//------------------------------------------------------------------------------
// HMI : input registers (1001...), REAL = low word first
//------------------------------------------------------------------------------
	//--- ADM100W_1
	GVL_MODBUS.Input_register_TCP_HMI[1000] := GVL_COM.COM_ADM100W_1.HMI_OUTPUT_FREQUENCY.Word_value[0];                   // 1001 | ADM100W Frequency (low word)
	GVL_MODBUS.Input_register_TCP_HMI[1001] := GVL_COM.COM_ADM100W_1.HMI_OUTPUT_FREQUENCY.Word_value[1];                   // 1002 | ADM100W Frequency (high word)
	GVL_MODBUS.Input_register_TCP_HMI[1002] := GVL_COM.COM_ADM100W_1.HMI_OUTPUT_L1_L2_VOLTAGE.Word_value[0];               // 1003 | ADM100W L1-L2 Voltage (low word)
	GVL_MODBUS.Input_register_TCP_HMI[1003] := GVL_COM.COM_ADM100W_1.HMI_OUTPUT_L1_L2_VOLTAGE.Word_value[1];               // 1004 | ADM100W L1-L2 Voltage (high word)
	GVL_MODBUS.Input_register_TCP_HMI[1004] := GVL_COM.COM_ADM100W_1.HMI_OUTPUT_L1_N_VOLTAGE.Word_value[0];                // 1005 | ADM100W L1-N Voltage (low word)
	GVL_MODBUS.Input_register_TCP_HMI[1005] := GVL_COM.COM_ADM100W_1.HMI_OUTPUT_L1_N_VOLTAGE.Word_value[1];                // 1006 | ADM100W L1-N Voltage (high word)
	GVL_MODBUS.Input_register_TCP_HMI[1006] := GVL_COM.COM_ADM100W_1.HMI_OUTPUT_L1_CURRENT.Word_value[0];                  // 1007 | ADM100W L1 Current (low word)
	GVL_MODBUS.Input_register_TCP_HMI[1007] := GVL_COM.COM_ADM100W_1.HMI_OUTPUT_L1_CURRENT.Word_value[1];                  // 1008 | ADM100W L1 Current (high word)
	GVL_MODBUS.Input_register_TCP_HMI[1008] := GVL_COM.COM_ADM100W_1.HMI_OUTPUT_L1_ACTIVE_POWER.Word_value[0];             // 1009 | ADM100W L1 Active Power (low word)
	GVL_MODBUS.Input_register_TCP_HMI[1009] := GVL_COM.COM_ADM100W_1.HMI_OUTPUT_L1_ACTIVE_POWER.Word_value[1];             // 1010 | ADM100W L1 Active Power (high word)
	GVL_MODBUS.Input_register_TCP_HMI[1010] := GVL_COM.COM_ADM100W_1.HMI_OUTPUT_L1_APPARENT_POWER.Word_value[0];           // 1011 | ADM100W L1 Apparent Power (low word)
	GVL_MODBUS.Input_register_TCP_HMI[1011] := GVL_COM.COM_ADM100W_1.HMI_OUTPUT_L1_APPARENT_POWER.Word_value[1];           // 1012 | ADM100W L1 Apparent Power (high word)
	GVL_MODBUS.Input_register_TCP_HMI[1012] := GVL_COM.COM_ADM100W_1.HMI_OUTPUT_L1_REACTIVE_POWER.Word_value[0];           // 1013 | ADM100W L1 Reactive Power (low word)
	GVL_MODBUS.Input_register_TCP_HMI[1013] := GVL_COM.COM_ADM100W_1.HMI_OUTPUT_L1_REACTIVE_POWER.Word_value[1];           // 1014 | ADM100W L1 Reactive Power (high word)
	GVL_MODBUS.Input_register_TCP_HMI[1014] := GVL_COM.COM_ADM100W_1.HMI_OUTPUT_L1_CURRENT_PHASE_ANGLE.Word_value[0];      // 1015 | ADM100W L1 Current Phase Angle (low word)
	GVL_MODBUS.Input_register_TCP_HMI[1015] := GVL_COM.COM_ADM100W_1.HMI_OUTPUT_L1_CURRENT_PHASE_ANGLE.Word_value[1];      // 1016 | ADM100W L1 Current Phase Angle (high word)
	GVL_MODBUS.Input_register_TCP_HMI[1016] := GVL_COM.COM_ADM100W_1.HMI_OUTPUT_L1_POWER_FACTOR.Word_value[0];             // 1017 | ADM100W L1 Power Factor (low word)
	GVL_MODBUS.Input_register_TCP_HMI[1017] := GVL_COM.COM_ADM100W_1.HMI_OUTPUT_L1_POWER_FACTOR.Word_value[1];             // 1018 | ADM100W L1 Power Factor (high word)
	GVL_MODBUS.Input_register_TCP_HMI[1018] := GVL_COM.COM_ADM100W_1.HMI_OUTPUT_L1_VOLTAGE_THD.Word_value[0];              // 1019 | ADM100W L1 Voltage THD (low word)
	GVL_MODBUS.Input_register_TCP_HMI[1019] := GVL_COM.COM_ADM100W_1.HMI_OUTPUT_L1_VOLTAGE_THD.Word_value[1];              // 1020 | ADM100W L1 Voltage THD (high word)
	GVL_MODBUS.Input_register_TCP_HMI[1020] := GVL_COM.COM_ADM100W_1.HMI_OUTPUT_L1_CURRENT_THD.Word_value[0];              // 1021 | ADM100W L1 Current THD (low word)
	GVL_MODBUS.Input_register_TCP_HMI[1021] := GVL_COM.COM_ADM100W_1.HMI_OUTPUT_L1_CURRENT_THD.Word_value[1];              // 1022 | ADM100W L1 Current THD (high word)
	GVL_MODBUS.Input_register_TCP_HMI[1022] := GVL_COM.COM_ADM100W_1.HMI_OUTPUT_L1_MAX_LOAD.Word_value[0];                 // 1023 | ADM100W L1 Max Load (low word)
	GVL_MODBUS.Input_register_TCP_HMI[1023] := GVL_COM.COM_ADM100W_1.HMI_OUTPUT_L1_MAX_LOAD.Word_value[1];                 // 1024 | ADM100W L1 Max Load (high word)
	GVL_MODBUS.Input_register_TCP_HMI[1024] := GVL_COM.COM_ADM100W_1.HMI_OUTPUT_L1_L2_VOLTAGE_PHASE_ANGLE.Word_value[0];   // 1025 | ADM100W L1-L2 Voltage Phase Angle (low word)
	GVL_MODBUS.Input_register_TCP_HMI[1025] := GVL_COM.COM_ADM100W_1.HMI_OUTPUT_L1_L2_VOLTAGE_PHASE_ANGLE.Word_value[1];   // 1026 | ADM100W L1-L2 Voltage Phase Angle (high word)
	GVL_MODBUS.Input_register_TCP_HMI[1026] := GVL_COM.COM_ADM100W_1.HMI_OUTPUT_L2_L3_VOLTAGE.Word_value[0];               // 1027 | ADM100W L2-L3 Voltage (low word)
	GVL_MODBUS.Input_register_TCP_HMI[1027] := GVL_COM.COM_ADM100W_1.HMI_OUTPUT_L2_L3_VOLTAGE.Word_value[1];               // 1028 | ADM100W L2-L3 Voltage (high word)
	GVL_MODBUS.Input_register_TCP_HMI[1028] := GVL_COM.COM_ADM100W_1.HMI_OUTPUT_L2_N_VOLTAGE.Word_value[0];                // 1029 | ADM100W L2-N Voltage (low word)
	GVL_MODBUS.Input_register_TCP_HMI[1029] := GVL_COM.COM_ADM100W_1.HMI_OUTPUT_L2_N_VOLTAGE.Word_value[1];                // 1030 | ADM100W L2-N Voltage (high word)
	GVL_MODBUS.Input_register_TCP_HMI[1030] := GVL_COM.COM_ADM100W_1.HMI_OUTPUT_L2_CURRENT.Word_value[0];                  // 1031 | ADM100W L2 Current (low word)
	GVL_MODBUS.Input_register_TCP_HMI[1031] := GVL_COM.COM_ADM100W_1.HMI_OUTPUT_L2_CURRENT.Word_value[1];                  // 1032 | ADM100W L2 Current (high word)
	GVL_MODBUS.Input_register_TCP_HMI[1032] := GVL_COM.COM_ADM100W_1.HMI_OUTPUT_L2_ACTIVE_POWER.Word_value[0];             // 1033 | ADM100W L2 Active Power (low word)
	GVL_MODBUS.Input_register_TCP_HMI[1033] := GVL_COM.COM_ADM100W_1.HMI_OUTPUT_L2_ACTIVE_POWER.Word_value[1];             // 1034 | ADM100W L2 Active Power (high word)
	GVL_MODBUS.Input_register_TCP_HMI[1034] := GVL_COM.COM_ADM100W_1.HMI_OUTPUT_L2_APPARENT_POWER.Word_value[0];           // 1035 | ADM100W L2 Apparent Power (low word)
	GVL_MODBUS.Input_register_TCP_HMI[1035] := GVL_COM.COM_ADM100W_1.HMI_OUTPUT_L2_APPARENT_POWER.Word_value[1];           // 1036 | ADM100W L2 Apparent Power (high word)
	GVL_MODBUS.Input_register_TCP_HMI[1036] := GVL_COM.COM_ADM100W_1.HMI_OUTPUT_L2_REACTIVE_POWER.Word_value[0];           // 1037 | ADM100W L2 Reactive Power (low word)
	GVL_MODBUS.Input_register_TCP_HMI[1037] := GVL_COM.COM_ADM100W_1.HMI_OUTPUT_L2_REACTIVE_POWER.Word_value[1];           // 1038 | ADM100W L2 Reactive Power (high word)
	GVL_MODBUS.Input_register_TCP_HMI[1038] := GVL_COM.COM_ADM100W_1.HMI_OUTPUT_L2_CURRENT_PHASE_ANGLE.Word_value[0];      // 1039 | ADM100W L2 Current Phase Angle (low word)
	GVL_MODBUS.Input_register_TCP_HMI[1039] := GVL_COM.COM_ADM100W_1.HMI_OUTPUT_L2_CURRENT_PHASE_ANGLE.Word_value[1];      // 1040 | ADM100W L2 Current Phase Angle (high word)
	GVL_MODBUS.Input_register_TCP_HMI[1040] := GVL_COM.COM_ADM100W_1.HMI_OUTPUT_L2_POWER_FACTOR.Word_value[0];             // 1041 | ADM100W L2 Power Factor (low word)
	GVL_MODBUS.Input_register_TCP_HMI[1041] := GVL_COM.COM_ADM100W_1.HMI_OUTPUT_L2_POWER_FACTOR.Word_value[1];             // 1042 | ADM100W L2 Power Factor (high word)
	GVL_MODBUS.Input_register_TCP_HMI[1042] := GVL_COM.COM_ADM100W_1.HMI_OUTPUT_L2_VOLTAGE_THD.Word_value[0];              // 1043 | ADM100W L2 Voltage THD (low word)
	GVL_MODBUS.Input_register_TCP_HMI[1043] := GVL_COM.COM_ADM100W_1.HMI_OUTPUT_L2_VOLTAGE_THD.Word_value[1];              // 1044 | ADM100W L2 Voltage THD (high word)
	GVL_MODBUS.Input_register_TCP_HMI[1044] := GVL_COM.COM_ADM100W_1.HMI_OUTPUT_L2_CURRENT_THD.Word_value[0];              // 1045 | ADM100W L2 Current THD (low word)
	GVL_MODBUS.Input_register_TCP_HMI[1045] := GVL_COM.COM_ADM100W_1.HMI_OUTPUT_L2_CURRENT_THD.Word_value[1];              // 1046 | ADM100W L2 Current THD (high word)
	GVL_MODBUS.Input_register_TCP_HMI[1046] := GVL_COM.COM_ADM100W_1.HMI_OUTPUT_L2_MAX_LOAD.Word_value[0];                 // 1047 | ADM100W L2 Max Load (low word)
	GVL_MODBUS.Input_register_TCP_HMI[1047] := GVL_COM.COM_ADM100W_1.HMI_OUTPUT_L2_MAX_LOAD.Word_value[1];                 // 1048 | ADM100W L2 Max Load (high word)
	GVL_MODBUS.Input_register_TCP_HMI[1048] := GVL_COM.COM_ADM100W_1.HMI_OUTPUT_L1_L3_VOLTAGE_PHASE_ANGLE.Word_value[0];   // 1049 | ADM100W L1-L3 Voltage Phase Angle (low word)
	GVL_MODBUS.Input_register_TCP_HMI[1049] := GVL_COM.COM_ADM100W_1.HMI_OUTPUT_L1_L3_VOLTAGE_PHASE_ANGLE.Word_value[1];   // 1050 | ADM100W L1-L3 Voltage Phase Angle (high word)
	GVL_MODBUS.Input_register_TCP_HMI[1050] := GVL_COM.COM_ADM100W_1.HMI_OUTPUT_L3_L1_VOLTAGE.Word_value[0];               // 1051 | ADM100W L3-L1 Voltage (low word)
	GVL_MODBUS.Input_register_TCP_HMI[1051] := GVL_COM.COM_ADM100W_1.HMI_OUTPUT_L3_L1_VOLTAGE.Word_value[1];               // 1052 | ADM100W L3-L1 Voltage (high word)
	GVL_MODBUS.Input_register_TCP_HMI[1052] := GVL_COM.COM_ADM100W_1.HMI_OUTPUT_L3_N_VOLTAGE.Word_value[0];                // 1053 | ADM100W L3-N Voltage (low word)
	GVL_MODBUS.Input_register_TCP_HMI[1053] := GVL_COM.COM_ADM100W_1.HMI_OUTPUT_L3_N_VOLTAGE.Word_value[1];                // 1054 | ADM100W L3-N Voltage (high word)
	GVL_MODBUS.Input_register_TCP_HMI[1054] := GVL_COM.COM_ADM100W_1.HMI_OUTPUT_L3_CURRENT.Word_value[0];                  // 1055 | ADM100W L3 Current (low word)
	GVL_MODBUS.Input_register_TCP_HMI[1055] := GVL_COM.COM_ADM100W_1.HMI_OUTPUT_L3_CURRENT.Word_value[1];                  // 1056 | ADM100W L3 Current (high word)
	GVL_MODBUS.Input_register_TCP_HMI[1056] := GVL_COM.COM_ADM100W_1.HMI_OUTPUT_L3_ACTIVE_POWER.Word_value[0];             // 1057 | ADM100W L3 Active Power (low word)
	GVL_MODBUS.Input_register_TCP_HMI[1057] := GVL_COM.COM_ADM100W_1.HMI_OUTPUT_L3_ACTIVE_POWER.Word_value[1];             // 1058 | ADM100W L3 Active Power (high word)
	GVL_MODBUS.Input_register_TCP_HMI[1058] := GVL_COM.COM_ADM100W_1.HMI_OUTPUT_L3_APPARENT_POWER.Word_value[0];           // 1059 | ADM100W L3 Apparent Power (low word)
	GVL_MODBUS.Input_register_TCP_HMI[1059] := GVL_COM.COM_ADM100W_1.HMI_OUTPUT_L3_APPARENT_POWER.Word_value[1];           // 1060 | ADM100W L3 Apparent Power (high word)
	GVL_MODBUS.Input_register_TCP_HMI[1060] := GVL_COM.COM_ADM100W_1.HMI_OUTPUT_L3_REACTIVE_POWER.Word_value[0];           // 1061 | ADM100W L3 Reactive Power (low word)
	GVL_MODBUS.Input_register_TCP_HMI[1061] := GVL_COM.COM_ADM100W_1.HMI_OUTPUT_L3_REACTIVE_POWER.Word_value[1];           // 1062 | ADM100W L3 Reactive Power (high word)
	GVL_MODBUS.Input_register_TCP_HMI[1062] := GVL_COM.COM_ADM100W_1.HMI_OUTPUT_L3_CURRENT_PHASE_ANGLE.Word_value[0];      // 1063 | ADM100W L3 Current Phase Angle (low word)
	GVL_MODBUS.Input_register_TCP_HMI[1063] := GVL_COM.COM_ADM100W_1.HMI_OUTPUT_L3_CURRENT_PHASE_ANGLE.Word_value[1];      // 1064 | ADM100W L3 Current Phase Angle (high word)
	GVL_MODBUS.Input_register_TCP_HMI[1064] := GVL_COM.COM_ADM100W_1.HMI_OUTPUT_L3_POWER_FACTOR.Word_value[0];             // 1065 | ADM100W L3 Power Factor (low word)
	GVL_MODBUS.Input_register_TCP_HMI[1065] := GVL_COM.COM_ADM100W_1.HMI_OUTPUT_L3_POWER_FACTOR.Word_value[1];             // 1066 | ADM100W L3 Power Factor (high word)
	GVL_MODBUS.Input_register_TCP_HMI[1066] := GVL_COM.COM_ADM100W_1.HMI_OUTPUT_L3_VOLTAGE_THD.Word_value[0];              // 1067 | ADM100W L3 Voltage THD (low word)
	GVL_MODBUS.Input_register_TCP_HMI[1067] := GVL_COM.COM_ADM100W_1.HMI_OUTPUT_L3_VOLTAGE_THD.Word_value[1];              // 1068 | ADM100W L3 Voltage THD (high word)
	GVL_MODBUS.Input_register_TCP_HMI[1068] := GVL_COM.COM_ADM100W_1.HMI_OUTPUT_L3_CURRENT_THD.Word_value[0];              // 1069 | ADM100W L3 Current THD (low word)
	GVL_MODBUS.Input_register_TCP_HMI[1069] := GVL_COM.COM_ADM100W_1.HMI_OUTPUT_L3_CURRENT_THD.Word_value[1];              // 1070 | ADM100W L3 Current THD (high word)
	GVL_MODBUS.Input_register_TCP_HMI[1070] := GVL_COM.COM_ADM100W_1.HMI_OUTPUT_L3_MAX_LOAD.Word_value[0];                 // 1071 | ADM100W L3 Max Load (low word)
	GVL_MODBUS.Input_register_TCP_HMI[1071] := GVL_COM.COM_ADM100W_1.HMI_OUTPUT_L3_MAX_LOAD.Word_value[1];                 // 1072 | ADM100W L3 Max Load (high word)
	GVL_MODBUS.Input_register_TCP_HMI[1072] := GVL_COM.COM_ADM100W_1.HMI_OUTPUT_INTERNAL_TEMPERATURE.Word_value[0];        // 1073 | ADM100W Internal Temperature (low word)
	GVL_MODBUS.Input_register_TCP_HMI[1073] := GVL_COM.COM_ADM100W_1.HMI_OUTPUT_INTERNAL_TEMPERATURE.Word_value[1];        // 1074 | ADM100W Internal Temperature (high word)
	GVL_MODBUS.Input_register_TCP_HMI[1074] := GVL_COM.COM_ADM100W_1.HMI_OUTPUT_ACTIVE_ENERGY.Word_value[0];               // 1075 | ADM100W Active Energy (low word)
	GVL_MODBUS.Input_register_TCP_HMI[1075] := GVL_COM.COM_ADM100W_1.HMI_OUTPUT_ACTIVE_ENERGY.Word_value[1];               // 1076 | ADM100W Active Energy (high word)
	GVL_MODBUS.Input_register_TCP_HMI[1076] := GVL_COM.COM_ADM100W_1.HMI_OUTPUT_APPARENT_ENERGY.Word_value[0];             // 1077 | ADM100W Apparent Energy (low word)
	GVL_MODBUS.Input_register_TCP_HMI[1077] := GVL_COM.COM_ADM100W_1.HMI_OUTPUT_APPARENT_ENERGY.Word_value[1];             // 1078 | ADM100W Apparent Energy (high word)
	GVL_MODBUS.Input_register_TCP_HMI[1078] := GVL_COM.COM_ADM100W_1.HMI_OUTPUT_REACTIVE_ENERGY.Word_value[0];             // 1079 | ADM100W Reactive Energy (low word)
	GVL_MODBUS.Input_register_TCP_HMI[1079] := GVL_COM.COM_ADM100W_1.HMI_OUTPUT_REACTIVE_ENERGY.Word_value[1];             // 1080 | ADM100W Reactive Energy (high word)
	GVL_MODBUS.Input_register_TCP_HMI[1080] := GVL_COM.COM_ADM100W_1.HMI_OUTPUT_TOTAL_ACTIVE_POWER.Word_value[0];          // 1081 | ADM100W Total Active Power (low word)
	GVL_MODBUS.Input_register_TCP_HMI[1081] := GVL_COM.COM_ADM100W_1.HMI_OUTPUT_TOTAL_ACTIVE_POWER.Word_value[1];          // 1082 | ADM100W Total Active Power (high word)
	GVL_MODBUS.Input_register_TCP_HMI[1082] := GVL_COM.COM_ADM100W_1.HMI_OUTPUT_TOTAL_APPARENT_POWER.Word_value[0];        // 1083 | ADM100W Total Apparent Power (low word)
	GVL_MODBUS.Input_register_TCP_HMI[1083] := GVL_COM.COM_ADM100W_1.HMI_OUTPUT_TOTAL_APPARENT_POWER.Word_value[1];        // 1084 | ADM100W Total Apparent Power (high word)
	GVL_MODBUS.Input_register_TCP_HMI[1084] := GVL_COM.COM_ADM100W_1.HMI_OUTPUT_TOTAL_REACTIVE_POWER.Word_value[0];        // 1085 | ADM100W Total Reactive Power (low word)
	GVL_MODBUS.Input_register_TCP_HMI[1085] := GVL_COM.COM_ADM100W_1.HMI_OUTPUT_TOTAL_REACTIVE_POWER.Word_value[1];        // 1086 | ADM100W Total Reactive Power (high word)
	GVL_MODBUS.Input_register_TCP_HMI[1086] := GVL_COM.COM_ADM100W_1.HMI_OUTPUT_ALL_PHASE_POWER_FACTOR.Word_value[0];      // 1087 | ADM100W All Phase Power Factor (low word)
	GVL_MODBUS.Input_register_TCP_HMI[1087] := GVL_COM.COM_ADM100W_1.HMI_OUTPUT_ALL_PHASE_POWER_FACTOR.Word_value[1];      // 1088 | ADM100W All Phase Power Factor (high word)

	//--- DOSENSOR_1
	GVL_MODBUS.Input_register_TCP_HMI[1088] := GVL_COM.COM_DOSENSOR_1.HMI_OUTPUT_SIGNAL.Word_value[0];   // 1089 | DO Sensor Signal (low word)
	GVL_MODBUS.Input_register_TCP_HMI[1089] := GVL_COM.COM_DOSENSOR_1.HMI_OUTPUT_SIGNAL.Word_value[1];   // 1090 | DO Sensor Signal (high word)

	//--- DIP1500_1
	GVL_MODBUS.Input_register_TCP_HMI[1090] := GVL_COM.COM_DIP1500_1.HMI_OUTPUT_FIRMWARE_VERSION;                               // 1091 | DIP1500 Firmware Version
	GVL_MODBUS.Input_register_TCP_HMI[1091] := GVL_COM.COM_DIP1500_1.HMI_OUTPUT_HARDWARE_VERSION;                               // 1092 | DIP1500 Hardware Version
	GVL_MODBUS.Input_register_TCP_HMI[1092] := GVL_COM.COM_DIP1500_1.HMI_OUTPUT_TEMPERATURE;                                    // 1093 | DIP1500 Temperature
	GVL_MODBUS.Input_register_TCP_HMI[1093] := GVL_COM.COM_DIP1500_1.HMI_OUTPUT_FLOAT_LEVEL_ALARM;                              // 1094 | DIP1500 Float Level Alarm
	GVL_MODBUS.Input_register_TCP_HMI[1094] := GVL_COM.COM_DIP1500_1.HMI_OUTPUT_DIGITAL_OUTPUT_VALUE;                           // 1095 | DIP1500 Digital Output Value
	GVL_MODBUS.Input_register_TCP_HMI[1095] := GVL_COM.COM_DIP1500_1.HMI_OUTPUT_REAL_TIME_RUN_TIME_OR_VOLUME.Word_value[0];     // 1096 | DIP1500 Real-Time Run Time Or Volume (low word)
	GVL_MODBUS.Input_register_TCP_HMI[1096] := GVL_COM.COM_DIP1500_1.HMI_OUTPUT_REAL_TIME_RUN_TIME_OR_VOLUME.Word_value[1];     // 1097 | DIP1500 Real-Time Run Time Or Volume (high word)
	GVL_MODBUS.Input_register_TCP_HMI[1097] := GVL_COM.COM_DIP1500_1.HMI_OUTPUT_ACCUMULATED_RUN_TIME_OR_VOLUME.Word_value[0];   // 1098 | DIP1500 Accumulated Run Time Or Volume (low word)
	GVL_MODBUS.Input_register_TCP_HMI[1098] := GVL_COM.COM_DIP1500_1.HMI_OUTPUT_ACCUMULATED_RUN_TIME_OR_VOLUME.Word_value[1];   // 1099 | DIP1500 Accumulated Run Time Or Volume (high word)

GFC_COM_OUT := TRUE;

          
END_FUNCTION

FUNCTION GFC_EXC_IN : BOOL

            
//==============================================================================
// GFC_EXC_IN
// GVL_EXC -> GVL_EXC : functional units (UPI) to equipment, before GFB_INST
// Simple copies only, no conversion (conversions are done in the FBs)
//==============================================================================

//------------------------------------------------------------------------------
// Global local modes (UPI_LOCAL_FUXA, UPI_LOCAL_HMI, UPI_LOCAL_WEBVISU) to every equipment
//------------------------------------------------------------------------------
	//--- ADM100W_1
	GVL_EXC.EXC_ADM100W_1.UPI_INPUT_GLOBAL_LOCAL_FUXA := GVL_EXC.EXC_UPI_LOCAL_FUXA.UPI_OUTPUT_LOCAL_ACTIVE;
	GVL_EXC.EXC_ADM100W_1.UPI_INPUT_GLOBAL_LOCAL_HMI  := GVL_EXC.EXC_UPI_LOCAL_HMI.UPI_OUTPUT_LOCAL_ACTIVE;
	GVL_EXC.EXC_ADM100W_1.UPI_INPUT_GLOBAL_LOCAL_WEBVISU := GVL_EXC.EXC_UPI_LOCAL_WEBVISU.UPI_OUTPUT_LOCAL_ACTIVE;

	//--- DOSENSOR_1
	GVL_EXC.EXC_DOSENSOR_1.UPI_INPUT_GLOBAL_LOCAL_FUXA := GVL_EXC.EXC_UPI_LOCAL_FUXA.UPI_OUTPUT_LOCAL_ACTIVE;
	GVL_EXC.EXC_DOSENSOR_1.UPI_INPUT_GLOBAL_LOCAL_HMI  := GVL_EXC.EXC_UPI_LOCAL_HMI.UPI_OUTPUT_LOCAL_ACTIVE;
	GVL_EXC.EXC_DOSENSOR_1.UPI_INPUT_GLOBAL_LOCAL_WEBVISU := GVL_EXC.EXC_UPI_LOCAL_WEBVISU.UPI_OUTPUT_LOCAL_ACTIVE;

	//--- DIP1500_1
	GVL_EXC.EXC_DIP1500_1.UPI_INPUT_GLOBAL_LOCAL_FUXA := GVL_EXC.EXC_UPI_LOCAL_FUXA.UPI_OUTPUT_LOCAL_ACTIVE;
	GVL_EXC.EXC_DIP1500_1.UPI_INPUT_GLOBAL_LOCAL_HMI  := GVL_EXC.EXC_UPI_LOCAL_HMI.UPI_OUTPUT_LOCAL_ACTIVE;
	GVL_EXC.EXC_DIP1500_1.UPI_INPUT_GLOBAL_LOCAL_WEBVISU := GVL_EXC.EXC_UPI_LOCAL_WEBVISU.UPI_OUTPUT_LOCAL_ACTIVE;

GFC_EXC_IN := TRUE;

          
END_FUNCTION

FUNCTION GFC_EXC_OUT : BOOL

            
//==============================================================================
// GFC_EXC_OUT
// GVL_EXC -> GVL_EXC : equipment to equipment, after GFB_INST
// Simple copies only, no conversion (conversions are done in the FBs)
//==============================================================================

// Nothing to copy yet
GFC_EXC_OUT := TRUE;

          
END_FUNCTION

FUNCTION GFC_IO_IN : BOOL

            
//==============================================================================
// GFC_IO_IN
// GVL_IOMAP (PLC I/O cards) -> GVL_IO
// Simple copies only, no conversion (conversions are done in the FBs)
//==============================================================================

//------------------------------------------------------------------------------
// Digital inputs
//------------------------------------------------------------------------------
	//--- DOSENSOR_1
	GVL_IO.IO_DOSENSOR_1.INPUT_SENSOR_FAULT := GVL_IOMAP.IOMAP_DI_FAULT_DOSENSOR_1;


//------------------------------------------------------------------------------
// Analog inputs
//------------------------------------------------------------------------------
	//--- DOSENSOR_1
	GVL_IO.IO_DOSENSOR_1.INPUT_SIGNAL := GVL_IOMAP.IOMAP_AI_SIGNAL_DOSENSOR_1;

GFC_IO_IN := TRUE;

          
END_FUNCTION

FUNCTION GFC_IO_OUT : BOOL

            
//==============================================================================
// GFC_IO_OUT
// GVL_IO -> GVL_IOMAP (PLC I/O cards)
// Simple copies only, no conversion (conversions are done in the FBs)
//==============================================================================

//------------------------------------------------------------------------------
// Digital outputs
//------------------------------------------------------------------------------
	//--- DOSENSOR_1
	GVL_IOMAP.IOMAP_DO_HIGH_DOSENSOR_1 := GVL_IO.IO_DOSENSOR_1.OUTPUT_CALIBRATION_HIGH;
	GVL_IOMAP.IOMAP_DO_LOW_DOSENSOR_1  := GVL_IO.IO_DOSENSOR_1.OUTPUT_CALIBRATION_LOW;

GFC_IO_OUT := TRUE;

          
END_FUNCTION

FUNCTION_BLOCK FB_UPI_LOCAL_FUXA
  VAR_IN_OUT
    COM : DUT_COM_UPI_LOCAL_FUXA;  (* Requests and status with SCADA / HMI *)
    EXC : DUT_EXC_UPI_LOCAL_FUXA;  (* Status to equipment *)
  END_VAR
  VAR
    INTERN : DUT_INT_UPI_LOCAL_FUXA;  (* Internal variables *)
  END_VAR

            
//==============================================================================
// FB_UPI_LOCAL_FUXA
// Global FUXA local mode for every equipment
// Set by the FUXA local request, reset by the FUXA auto request (pulse or maintained, auto wins)
// The equipment read this status through GFC_EXC_IN and report their own local status themselves
//==============================================================================

//------------------------------------------------------------------------------
// 1. INPUTS
//------------------------------------------------------------------------------
	INTERN.LOCAL_REQUEST := COM.SCADA_INPUT_LOCAL_REQUEST;
	INTERN.AUTO_REQUEST  := COM.SCADA_INPUT_AUTO_REQUEST;


//------------------------------------------------------------------------------
// 2. PROCESSING
//------------------------------------------------------------------------------
	IF INTERN.LOCAL_REQUEST THEN
		INTERN.LOCAL_ACTIVE := TRUE;
	END_IF
	IF INTERN.AUTO_REQUEST THEN
		INTERN.LOCAL_ACTIVE := FALSE;
	END_IF


//------------------------------------------------------------------------------
// 3. OUTPUTS
//------------------------------------------------------------------------------
	//--- EXC : to every equipment (through GFC_EXC_IN)
	EXC.UPI_OUTPUT_LOCAL_ACTIVE := INTERN.LOCAL_ACTIVE;

	//--- COM : status
	COM.SCADA_OUTPUT_LOCAL_ACTIVE := INTERN.LOCAL_ACTIVE;


          
END_FUNCTION_BLOCK

FUNCTION_BLOCK FB_UPI_LOCAL_HMI
  VAR_IN_OUT
    COM : DUT_COM_UPI_LOCAL_HMI;  (* Requests and status with SCADA / HMI *)
    EXC : DUT_EXC_UPI_LOCAL_HMI;  (* Status to equipment *)
  END_VAR
  VAR
    INTERN : DUT_INT_UPI_LOCAL_HMI;  (* Internal variables *)
  END_VAR

            
//==============================================================================
// FB_UPI_LOCAL_HMI
// Global HMI local mode for every equipment
// Set by the HMI local request, reset by the HMI auto request (pulse or maintained, auto wins)
// The equipment read this status through GFC_EXC_IN and report their own local status themselves
//==============================================================================

//------------------------------------------------------------------------------
// 1. INPUTS
//------------------------------------------------------------------------------
	INTERN.LOCAL_REQUEST := COM.HMI_INPUT_LOCAL_REQUEST;
	INTERN.AUTO_REQUEST  := COM.HMI_INPUT_AUTO_REQUEST;


//------------------------------------------------------------------------------
// 2. PROCESSING
//------------------------------------------------------------------------------
	IF INTERN.LOCAL_REQUEST THEN
		INTERN.LOCAL_ACTIVE := TRUE;
	END_IF
	IF INTERN.AUTO_REQUEST THEN
		INTERN.LOCAL_ACTIVE := FALSE;
	END_IF


//------------------------------------------------------------------------------
// 3. OUTPUTS
//------------------------------------------------------------------------------
	//--- EXC : to every equipment (through GFC_EXC_IN)
	EXC.UPI_OUTPUT_LOCAL_ACTIVE := INTERN.LOCAL_ACTIVE;

	//--- COM : status
	COM.HMI_OUTPUT_LOCAL_ACTIVE   := INTERN.LOCAL_ACTIVE;
	COM.SCADA_OUTPUT_LOCAL_ACTIVE := INTERN.LOCAL_ACTIVE;   // also reported to FUXA


          
END_FUNCTION_BLOCK

FUNCTION_BLOCK GFB_INST
  VAR
    FB_ADM100W_1 : FB_INST_ADM100W;  (* Trumeter ADM100W power meter *)
    FB_DOSENSOR_1 : FB_INST_DOSENSOR;  (* Dissolved oxygen sensor *)
    FB_DIP1500_1 : FB_INST_DIP1500;  (* Kamoer DIP1500 peristaltic pump *)
  END_VAR

            
//==============================================================================
// GFB_INST
// Calls every equipment instance
// One block per equipment, all interfaces connected
//==============================================================================

//--- ADM100W_1 : Trumeter ADM100W power meter
FB_ADM100W_1(
	PA  := GVL_PA.PA_ADM100W_1,
	COM := GVL_COM.COM_ADM100W_1,
	EXC := GVL_EXC.EXC_ADM100W_1,
	IO  := GVL_IO.IO_ADM100W_1);

//--- DOSENSOR_1 : Dissolved oxygen sensor
FB_DOSENSOR_1(
	PA  := GVL_PA.PA_DOSENSOR_1,
	COM := GVL_COM.COM_DOSENSOR_1,
	EXC := GVL_EXC.EXC_DOSENSOR_1,
	IO  := GVL_IO.IO_DOSENSOR_1);

//--- DIP1500_1 : Kamoer DIP1500 peristaltic pump
FB_DIP1500_1(
	PA  := GVL_PA.PA_DIP1500_1,
	COM := GVL_COM.COM_DIP1500_1,
	EXC := GVL_EXC.EXC_DIP1500_1,
	IO  := GVL_IO.IO_DIP1500_1);

          
END_FUNCTION_BLOCK

FUNCTION_BLOCK GFB_UPI
  VAR
    FB_UPI_LOCAL_FUXA_1 : FB_UPI_LOCAL_FUXA;  (* Global FUXA local mode *)
    FB_UPI_LOCAL_HMI_1 : FB_UPI_LOCAL_HMI;  (* Global HMI local mode *)
    FB_UPI_LOCAL_WEBVISU_1 : FB_UPI_LOCAL_WEBVISU;  (* Global WEBVISU local mode *)
  END_VAR

            
//==============================================================================
// GFB_UPI
// Calls every functional unit (UPI)
// Runs before GFB_INST, results go to the equipment through GFC_EXC_IN
//==============================================================================

//--- UPI_LOCAL_FUXA : Global FUXA local mode
FB_UPI_LOCAL_FUXA_1(
	COM := GVL_COM.COM_UPI_LOCAL_FUXA,
	EXC := GVL_EXC.EXC_UPI_LOCAL_FUXA);

//--- UPI_LOCAL_HMI : Global HMI local mode
FB_UPI_LOCAL_HMI_1(
	COM := GVL_COM.COM_UPI_LOCAL_HMI,
	EXC := GVL_EXC.EXC_UPI_LOCAL_HMI);

//--- UPI_LOCAL_WEBVISU : Global WEBVISU local mode (direct IEC variables)
FB_UPI_LOCAL_WEBVISU_1(
	COM := GVL_COM.COM_UPI_LOCAL_WEBVISU,
	EXC := GVL_EXC.EXC_UPI_LOCAL_WEBVISU);

          
END_FUNCTION_BLOCK

FUNCTION_BLOCK FB_UPI_LOCAL_WEBVISU
  VAR_IN_OUT
    COM : DUT_COM_UPI_LOCAL_WEBVISU;  (* Direct IEC requests and status with WEBVISU *)
    EXC : DUT_EXC_UPI_LOCAL_WEBVISU;  (* Status to equipment *)
  END_VAR
  VAR
    INTERN : DUT_INT_UPI_LOCAL_WEBVISU;  (* Internal variables *)
  END_VAR

            
//==============================================================================
// FB_UPI_LOCAL_WEBVISU
// Global WEBVISU local mode for every equipment
// Set by the WEBVISU local request, reset by the WEBVISU auto request (pulse or maintained, auto wins)
// The equipment read this status through GFC_EXC_IN and report their own local status themselves
//==============================================================================

//------------------------------------------------------------------------------
// 1. INPUTS
//------------------------------------------------------------------------------
	INTERN.LOCAL_REQUEST := COM.WEBVISU_INPUT_LOCAL_REQUEST;
	INTERN.AUTO_REQUEST  := COM.WEBVISU_INPUT_AUTO_REQUEST;


//------------------------------------------------------------------------------
// 2. PROCESSING
//------------------------------------------------------------------------------
	IF INTERN.LOCAL_REQUEST THEN
		INTERN.LOCAL_ACTIVE := TRUE;
	END_IF
	IF INTERN.AUTO_REQUEST THEN
		INTERN.LOCAL_ACTIVE := FALSE;
	END_IF


//------------------------------------------------------------------------------
// 3. OUTPUTS
//------------------------------------------------------------------------------
	//--- EXC : to every equipment (through GFC_EXC_IN)
	EXC.UPI_OUTPUT_LOCAL_ACTIVE := INTERN.LOCAL_ACTIVE;

	//--- COM : status
	COM.WEBVISU_OUTPUT_LOCAL_ACTIVE := INTERN.LOCAL_ACTIVE;


          
END_FUNCTION_BLOCK

FUNCTION_BLOCK FB_INST_ADM100W
  VAR_IN_OUT
    PA : DUT_PA_ADM100W;  (* Parameters (persistent, GVL_PA) *)
    COM : DUT_COM_ADM100W;  (* Communication : Modbus RTU (COM_), SCADA FUXA (SCADA_), HMI (HMI_) *)
    EXC : DUT_EXC_ADM100W;  (* Exchanges : other equipment (EXC_), functional units (UPI_) *)
    IO : DUT_IO_ADM100W;  (* Wired PLC I/O *)
  END_VAR
  VAR
    INTERN : DUT_INT_ADM100W;  (* Internal variables *)
  END_VAR

            
//==============================================================================
// FB_INST_ADM100W
// Trumeter ADM100W power meter, Modbus RTU, 32-bit float MSW first (ABCD). No command : local mode is only reported
// 1. INPUTS     : requests, control mode, command source, equipment feedback -> INTERN
// 2. PROCESSING : on INTERN only
// 3. OUTPUTS    : INTERN -> COM / IO / EXC
// Control mode  : local WEBVISU > local HMI > local FUXA > auto (functional units)
//==============================================================================

//------------------------------------------------------------------------------
// 1. INPUTS
//------------------------------------------------------------------------------
	//--- Control mode requests (WEBVISU, HMI, FUXA, global UPI)
	INTERN.FUXA_LOCAL_REQUEST := COM.SCADA_INPUT_LOCAL_REQUEST;
	INTERN.FUXA_AUTO_REQUEST  := COM.SCADA_INPUT_AUTO_REQUEST;
	INTERN.HMI_LOCAL_REQUEST  := COM.HMI_INPUT_LOCAL_REQUEST;
	INTERN.HMI_AUTO_REQUEST   := COM.HMI_INPUT_AUTO_REQUEST;
	INTERN.GLOBAL_LOCAL_FUXA  := EXC.UPI_INPUT_GLOBAL_LOCAL_FUXA;
	INTERN.GLOBAL_LOCAL_HMI   := EXC.UPI_INPUT_GLOBAL_LOCAL_HMI;
	INTERN.WEBVISU_LOCAL_REQUEST := COM.WEBVISU_INPUT_LOCAL_REQUEST;
	INTERN.WEBVISU_AUTO_REQUEST  := COM.WEBVISU_INPUT_AUTO_REQUEST;
	INTERN.GLOBAL_LOCAL_WEBVISU  := EXC.UPI_INPUT_GLOBAL_LOCAL_WEBVISU;

	//--- Control mode
	// Individual memories : set by the local request, reset by the auto request (auto wins if both)
	IF INTERN.WEBVISU_LOCAL_REQUEST THEN
		INTERN.LOCAL_WEBVISU_INDIVIDUAL := TRUE;
	END_IF
	IF INTERN.WEBVISU_AUTO_REQUEST THEN
		INTERN.LOCAL_WEBVISU_INDIVIDUAL := FALSE;
	END_IF
	IF INTERN.HMI_LOCAL_REQUEST THEN
		INTERN.LOCAL_HMI_INDIVIDUAL := TRUE;
	END_IF
	IF INTERN.HMI_AUTO_REQUEST THEN
		INTERN.LOCAL_HMI_INDIVIDUAL := FALSE;
	END_IF
	IF INTERN.FUXA_LOCAL_REQUEST THEN
		INTERN.LOCAL_FUXA_INDIVIDUAL := TRUE;
	END_IF
	IF INTERN.FUXA_AUTO_REQUEST THEN
		INTERN.LOCAL_FUXA_INDIVIDUAL := FALSE;
	END_IF

	// Resulting mode : individual OR global, WEBVISU > HMI > FUXA > auto
	INTERN.LOCAL_WEBVISU := INTERN.LOCAL_WEBVISU_INDIVIDUAL OR INTERN.GLOBAL_LOCAL_WEBVISU;
	INTERN.LOCAL_HMI     := (INTERN.LOCAL_HMI_INDIVIDUAL OR INTERN.GLOBAL_LOCAL_HMI) AND NOT INTERN.LOCAL_WEBVISU;
	INTERN.LOCAL_FUXA    := (INTERN.LOCAL_FUXA_INDIVIDUAL OR INTERN.GLOBAL_LOCAL_FUXA) AND NOT INTERN.LOCAL_WEBVISU AND NOT INTERN.LOCAL_HMI;
	INTERN.AUTO          := NOT INTERN.LOCAL_WEBVISU AND NOT INTERN.LOCAL_HMI AND NOT INTERN.LOCAL_FUXA;

	//--- COM : alarms (coils 0..9)
	INTERN.ALARM_1  := COM.COM_INPUT_COILS[0].0;
	INTERN.ALARM_2  := COM.COM_INPUT_COILS[0].1;
	INTERN.ALARM_3  := COM.COM_INPUT_COILS[0].2;
	INTERN.ALARM_4  := COM.COM_INPUT_COILS[0].3;
	INTERN.ALARM_5  := COM.COM_INPUT_COILS[0].4;
	INTERN.ALARM_6  := COM.COM_INPUT_COILS[0].5;
	INTERN.ALARM_7  := COM.COM_INPUT_COILS[0].6;
	INTERN.ALARM_8  := COM.COM_INPUT_COILS[0].7;
	INTERN.ALARM_9  := COM.COM_INPUT_COILS[1].0;
	INTERN.ALARM_10 := COM.COM_INPUT_COILS[1].1;

	//--- COM : measures (input registers, MSW first)
	INTERN.FREQUENCY                 := FNC_WORDS_TO_REAL(High_word := COM.COM_INPUT_IR[0], Low_word := COM.COM_INPUT_IR[1]);
	INTERN.L1_L2_VOLTAGE             := FNC_WORDS_TO_REAL(High_word := COM.COM_INPUT_IR[2], Low_word := COM.COM_INPUT_IR[3]);
	INTERN.L1_N_VOLTAGE              := FNC_WORDS_TO_REAL(High_word := COM.COM_INPUT_IR[4], Low_word := COM.COM_INPUT_IR[5]);
	INTERN.L1_CURRENT                := FNC_WORDS_TO_REAL(High_word := COM.COM_INPUT_IR[6], Low_word := COM.COM_INPUT_IR[7]);
	INTERN.L1_ACTIVE_POWER           := FNC_WORDS_TO_REAL(High_word := COM.COM_INPUT_IR[8], Low_word := COM.COM_INPUT_IR[9]);
	INTERN.L1_APPARENT_POWER         := FNC_WORDS_TO_REAL(High_word := COM.COM_INPUT_IR[10], Low_word := COM.COM_INPUT_IR[11]);
	INTERN.L1_REACTIVE_POWER         := FNC_WORDS_TO_REAL(High_word := COM.COM_INPUT_IR[12], Low_word := COM.COM_INPUT_IR[13]);
	INTERN.L1_CURRENT_PHASE_ANGLE    := FNC_WORDS_TO_REAL(High_word := COM.COM_INPUT_IR[14], Low_word := COM.COM_INPUT_IR[15]);
	INTERN.L1_POWER_FACTOR           := FNC_WORDS_TO_REAL(High_word := COM.COM_INPUT_IR[16], Low_word := COM.COM_INPUT_IR[17]);
	INTERN.L1_VOLTAGE_THD            := FNC_WORDS_TO_REAL(High_word := COM.COM_INPUT_IR[18], Low_word := COM.COM_INPUT_IR[19]);
	INTERN.L1_CURRENT_THD            := FNC_WORDS_TO_REAL(High_word := COM.COM_INPUT_IR[20], Low_word := COM.COM_INPUT_IR[21]);
	INTERN.L1_MAX_LOAD               := FNC_WORDS_TO_REAL(High_word := COM.COM_INPUT_IR[22], Low_word := COM.COM_INPUT_IR[23]);
	INTERN.L1_L2_VOLTAGE_PHASE_ANGLE := FNC_WORDS_TO_REAL(High_word := COM.COM_INPUT_IR[24], Low_word := COM.COM_INPUT_IR[25]);
	INTERN.L2_L3_VOLTAGE             := FNC_WORDS_TO_REAL(High_word := COM.COM_INPUT_IR[26], Low_word := COM.COM_INPUT_IR[27]);
	INTERN.L2_N_VOLTAGE              := FNC_WORDS_TO_REAL(High_word := COM.COM_INPUT_IR[28], Low_word := COM.COM_INPUT_IR[29]);
	INTERN.L2_CURRENT                := FNC_WORDS_TO_REAL(High_word := COM.COM_INPUT_IR[30], Low_word := COM.COM_INPUT_IR[31]);
	INTERN.L2_ACTIVE_POWER           := FNC_WORDS_TO_REAL(High_word := COM.COM_INPUT_IR[32], Low_word := COM.COM_INPUT_IR[33]);
	INTERN.L2_APPARENT_POWER         := FNC_WORDS_TO_REAL(High_word := COM.COM_INPUT_IR[34], Low_word := COM.COM_INPUT_IR[35]);
	INTERN.L2_REACTIVE_POWER         := FNC_WORDS_TO_REAL(High_word := COM.COM_INPUT_IR[36], Low_word := COM.COM_INPUT_IR[37]);
	INTERN.L2_CURRENT_PHASE_ANGLE    := FNC_WORDS_TO_REAL(High_word := COM.COM_INPUT_IR[38], Low_word := COM.COM_INPUT_IR[39]);
	INTERN.L2_POWER_FACTOR           := FNC_WORDS_TO_REAL(High_word := COM.COM_INPUT_IR[40], Low_word := COM.COM_INPUT_IR[41]);
	INTERN.L2_VOLTAGE_THD            := FNC_WORDS_TO_REAL(High_word := COM.COM_INPUT_IR[42], Low_word := COM.COM_INPUT_IR[43]);
	INTERN.L2_CURRENT_THD            := FNC_WORDS_TO_REAL(High_word := COM.COM_INPUT_IR[44], Low_word := COM.COM_INPUT_IR[45]);
	INTERN.L2_MAX_LOAD               := FNC_WORDS_TO_REAL(High_word := COM.COM_INPUT_IR[46], Low_word := COM.COM_INPUT_IR[47]);
	INTERN.L1_L3_VOLTAGE_PHASE_ANGLE := FNC_WORDS_TO_REAL(High_word := COM.COM_INPUT_IR[48], Low_word := COM.COM_INPUT_IR[49]);
	INTERN.L3_L1_VOLTAGE             := FNC_WORDS_TO_REAL(High_word := COM.COM_INPUT_IR[50], Low_word := COM.COM_INPUT_IR[51]);
	INTERN.L3_N_VOLTAGE              := FNC_WORDS_TO_REAL(High_word := COM.COM_INPUT_IR[52], Low_word := COM.COM_INPUT_IR[53]);
	INTERN.L3_CURRENT                := FNC_WORDS_TO_REAL(High_word := COM.COM_INPUT_IR[54], Low_word := COM.COM_INPUT_IR[55]);
	INTERN.L3_ACTIVE_POWER           := FNC_WORDS_TO_REAL(High_word := COM.COM_INPUT_IR[56], Low_word := COM.COM_INPUT_IR[57]);
	INTERN.L3_APPARENT_POWER         := FNC_WORDS_TO_REAL(High_word := COM.COM_INPUT_IR[58], Low_word := COM.COM_INPUT_IR[59]);
	INTERN.L3_REACTIVE_POWER         := FNC_WORDS_TO_REAL(High_word := COM.COM_INPUT_IR[60], Low_word := COM.COM_INPUT_IR[61]);
	INTERN.L3_CURRENT_PHASE_ANGLE    := FNC_WORDS_TO_REAL(High_word := COM.COM_INPUT_IR[62], Low_word := COM.COM_INPUT_IR[63]);
	INTERN.L3_POWER_FACTOR           := FNC_WORDS_TO_REAL(High_word := COM.COM_INPUT_IR[64], Low_word := COM.COM_INPUT_IR[65]);
	INTERN.L3_VOLTAGE_THD            := FNC_WORDS_TO_REAL(High_word := COM.COM_INPUT_IR[66], Low_word := COM.COM_INPUT_IR[67]);
	INTERN.L3_CURRENT_THD            := FNC_WORDS_TO_REAL(High_word := COM.COM_INPUT_IR[68], Low_word := COM.COM_INPUT_IR[69]);
	INTERN.L3_MAX_LOAD               := FNC_WORDS_TO_REAL(High_word := COM.COM_INPUT_IR[70], Low_word := COM.COM_INPUT_IR[71]);
	INTERN.INTERNAL_TEMPERATURE      := FNC_WORDS_TO_REAL(High_word := COM.COM_INPUT_IR[72], Low_word := COM.COM_INPUT_IR[73]);
	INTERN.ACTIVE_ENERGY             := FNC_WORDS_TO_REAL(High_word := COM.COM_INPUT_IR[74], Low_word := COM.COM_INPUT_IR[75]);
	INTERN.APPARENT_ENERGY           := FNC_WORDS_TO_REAL(High_word := COM.COM_INPUT_IR[76], Low_word := COM.COM_INPUT_IR[77]);
	INTERN.REACTIVE_ENERGY           := FNC_WORDS_TO_REAL(High_word := COM.COM_INPUT_IR[78], Low_word := COM.COM_INPUT_IR[79]);
	INTERN.TOTAL_ACTIVE_POWER        := FNC_WORDS_TO_REAL(High_word := COM.COM_INPUT_IR[80], Low_word := COM.COM_INPUT_IR[81]);
	INTERN.TOTAL_APPARENT_POWER      := FNC_WORDS_TO_REAL(High_word := COM.COM_INPUT_IR[82], Low_word := COM.COM_INPUT_IR[83]);
	INTERN.TOTAL_REACTIVE_POWER      := FNC_WORDS_TO_REAL(High_word := COM.COM_INPUT_IR[84], Low_word := COM.COM_INPUT_IR[85]);
	INTERN.ALL_PHASE_POWER_FACTOR    := FNC_WORDS_TO_REAL(High_word := COM.COM_INPUT_IR[86], Low_word := COM.COM_INPUT_IR[87]);


//------------------------------------------------------------------------------
// 2. PROCESSING
//------------------------------------------------------------------------------
	// Nothing


//------------------------------------------------------------------------------
// 3. OUTPUTS
//------------------------------------------------------------------------------
	//--- COM : control mode status to SCADA, HMI and WEBVISU
	COM.SCADA_OUTPUT_LOCAL_FUXA_ACTIVE := INTERN.LOCAL_FUXA;
	COM.SCADA_OUTPUT_LOCAL_HMI_ACTIVE  := INTERN.LOCAL_HMI;
	COM.HMI_OUTPUT_LOCAL_ACTIVE        := INTERN.LOCAL_HMI;
	COM.WEBVISU_OUTPUT_LOCAL_ACTIVE        := INTERN.LOCAL_WEBVISU;
	COM.WEBVISU_OUTPUT_LOCAL_HMI_ACTIVE  := INTERN.LOCAL_HMI;
	COM.WEBVISU_OUTPUT_LOCAL_FUXA_ACTIVE := INTERN.LOCAL_FUXA;

	//--- EXC
	EXC.EXC_OUTPUT_FREQUENCY            := INTERN.FREQUENCY;
	EXC.EXC_OUTPUT_L1_N_VOLTAGE         := INTERN.L1_N_VOLTAGE;
	EXC.EXC_OUTPUT_L1_CURRENT           := INTERN.L1_CURRENT;
	EXC.EXC_OUTPUT_L1_ACTIVE_POWER      := INTERN.L1_ACTIVE_POWER;
	EXC.EXC_OUTPUT_L1_APPARENT_POWER    := INTERN.L1_APPARENT_POWER;
	EXC.EXC_OUTPUT_L1_REACTIVE_POWER    := INTERN.L1_REACTIVE_POWER;
	EXC.EXC_OUTPUT_L1_POWER_FACTOR      := INTERN.L1_POWER_FACTOR;
	EXC.EXC_OUTPUT_L1_VOLTAGE_THD       := INTERN.L1_VOLTAGE_THD;
	EXC.EXC_OUTPUT_L1_CURRENT_THD       := INTERN.L1_CURRENT_THD;
	EXC.EXC_OUTPUT_L1_MAX_LOAD          := INTERN.L1_MAX_LOAD;
	EXC.EXC_OUTPUT_INTERNAL_TEMPERATURE := INTERN.INTERNAL_TEMPERATURE;
	EXC.EXC_OUTPUT_ACTIVE_ENERGY        := INTERN.ACTIVE_ENERGY;
	// EXC.EXC_OUTPUT_DATA_VALID : not managed yet (no Modbus diagnostic)

	//--- COM : alarms to SCADA, HMI and WEBVISU
	COM.SCADA_OUTPUT_ALARM_1_STATUS  := INTERN.ALARM_1;
	COM.HMI_OUTPUT_ALARM_1_STATUS    := INTERN.ALARM_1;
	COM.WEBVISU_OUTPUT_ALARM_1_STATUS    := INTERN.ALARM_1;
	COM.SCADA_OUTPUT_ALARM_2_STATUS  := INTERN.ALARM_2;
	COM.HMI_OUTPUT_ALARM_2_STATUS    := INTERN.ALARM_2;
	COM.WEBVISU_OUTPUT_ALARM_2_STATUS    := INTERN.ALARM_2;
	COM.SCADA_OUTPUT_ALARM_3_STATUS  := INTERN.ALARM_3;
	COM.HMI_OUTPUT_ALARM_3_STATUS    := INTERN.ALARM_3;
	COM.WEBVISU_OUTPUT_ALARM_3_STATUS    := INTERN.ALARM_3;
	COM.SCADA_OUTPUT_ALARM_4_STATUS  := INTERN.ALARM_4;
	COM.HMI_OUTPUT_ALARM_4_STATUS    := INTERN.ALARM_4;
	COM.WEBVISU_OUTPUT_ALARM_4_STATUS    := INTERN.ALARM_4;
	COM.SCADA_OUTPUT_ALARM_5_STATUS  := INTERN.ALARM_5;
	COM.HMI_OUTPUT_ALARM_5_STATUS    := INTERN.ALARM_5;
	COM.WEBVISU_OUTPUT_ALARM_5_STATUS    := INTERN.ALARM_5;
	COM.SCADA_OUTPUT_ALARM_6_STATUS  := INTERN.ALARM_6;
	COM.HMI_OUTPUT_ALARM_6_STATUS    := INTERN.ALARM_6;
	COM.WEBVISU_OUTPUT_ALARM_6_STATUS    := INTERN.ALARM_6;
	COM.SCADA_OUTPUT_ALARM_7_STATUS  := INTERN.ALARM_7;
	COM.HMI_OUTPUT_ALARM_7_STATUS    := INTERN.ALARM_7;
	COM.WEBVISU_OUTPUT_ALARM_7_STATUS    := INTERN.ALARM_7;
	COM.SCADA_OUTPUT_ALARM_8_STATUS  := INTERN.ALARM_8;
	COM.HMI_OUTPUT_ALARM_8_STATUS    := INTERN.ALARM_8;
	COM.WEBVISU_OUTPUT_ALARM_8_STATUS    := INTERN.ALARM_8;
	COM.SCADA_OUTPUT_ALARM_9_STATUS  := INTERN.ALARM_9;
	COM.HMI_OUTPUT_ALARM_9_STATUS    := INTERN.ALARM_9;
	COM.WEBVISU_OUTPUT_ALARM_9_STATUS    := INTERN.ALARM_9;
	COM.SCADA_OUTPUT_ALARM_10_STATUS := INTERN.ALARM_10;
	COM.HMI_OUTPUT_ALARM_10_STATUS   := INTERN.ALARM_10;
	COM.WEBVISU_OUTPUT_ALARM_10_STATUS   := INTERN.ALARM_10;

	//--- COM : measures to SCADA, HMI and WEBVISU
	COM.SCADA_OUTPUT_FREQUENCY.Real_value                 := INTERN.FREQUENCY;
	COM.HMI_OUTPUT_FREQUENCY.Real_value                   := INTERN.FREQUENCY;
	COM.WEBVISU_OUTPUT_FREQUENCY.Real_value                   := INTERN.FREQUENCY;
	COM.SCADA_OUTPUT_L1_L2_VOLTAGE.Real_value             := INTERN.L1_L2_VOLTAGE;
	COM.HMI_OUTPUT_L1_L2_VOLTAGE.Real_value               := INTERN.L1_L2_VOLTAGE;
	COM.WEBVISU_OUTPUT_L1_L2_VOLTAGE.Real_value               := INTERN.L1_L2_VOLTAGE;
	COM.SCADA_OUTPUT_L1_N_VOLTAGE.Real_value              := INTERN.L1_N_VOLTAGE;
	COM.HMI_OUTPUT_L1_N_VOLTAGE.Real_value                := INTERN.L1_N_VOLTAGE;
	COM.WEBVISU_OUTPUT_L1_N_VOLTAGE.Real_value                := INTERN.L1_N_VOLTAGE;
	COM.SCADA_OUTPUT_L1_CURRENT.Real_value                := INTERN.L1_CURRENT;
	COM.HMI_OUTPUT_L1_CURRENT.Real_value                  := INTERN.L1_CURRENT;
	COM.WEBVISU_OUTPUT_L1_CURRENT.Real_value                  := INTERN.L1_CURRENT;
	COM.SCADA_OUTPUT_L1_ACTIVE_POWER.Real_value           := INTERN.L1_ACTIVE_POWER;
	COM.HMI_OUTPUT_L1_ACTIVE_POWER.Real_value             := INTERN.L1_ACTIVE_POWER;
	COM.WEBVISU_OUTPUT_L1_ACTIVE_POWER.Real_value             := INTERN.L1_ACTIVE_POWER;
	COM.SCADA_OUTPUT_L1_APPARENT_POWER.Real_value         := INTERN.L1_APPARENT_POWER;
	COM.HMI_OUTPUT_L1_APPARENT_POWER.Real_value           := INTERN.L1_APPARENT_POWER;
	COM.WEBVISU_OUTPUT_L1_APPARENT_POWER.Real_value           := INTERN.L1_APPARENT_POWER;
	COM.SCADA_OUTPUT_L1_REACTIVE_POWER.Real_value         := INTERN.L1_REACTIVE_POWER;
	COM.HMI_OUTPUT_L1_REACTIVE_POWER.Real_value           := INTERN.L1_REACTIVE_POWER;
	COM.WEBVISU_OUTPUT_L1_REACTIVE_POWER.Real_value           := INTERN.L1_REACTIVE_POWER;
	COM.SCADA_OUTPUT_L1_CURRENT_PHASE_ANGLE.Real_value    := INTERN.L1_CURRENT_PHASE_ANGLE;
	COM.HMI_OUTPUT_L1_CURRENT_PHASE_ANGLE.Real_value      := INTERN.L1_CURRENT_PHASE_ANGLE;
	COM.WEBVISU_OUTPUT_L1_CURRENT_PHASE_ANGLE.Real_value      := INTERN.L1_CURRENT_PHASE_ANGLE;
	COM.SCADA_OUTPUT_L1_POWER_FACTOR.Real_value           := INTERN.L1_POWER_FACTOR;
	COM.HMI_OUTPUT_L1_POWER_FACTOR.Real_value             := INTERN.L1_POWER_FACTOR;
	COM.WEBVISU_OUTPUT_L1_POWER_FACTOR.Real_value             := INTERN.L1_POWER_FACTOR;
	COM.SCADA_OUTPUT_L1_VOLTAGE_THD.Real_value            := INTERN.L1_VOLTAGE_THD;
	COM.HMI_OUTPUT_L1_VOLTAGE_THD.Real_value              := INTERN.L1_VOLTAGE_THD;
	COM.WEBVISU_OUTPUT_L1_VOLTAGE_THD.Real_value              := INTERN.L1_VOLTAGE_THD;
	COM.SCADA_OUTPUT_L1_CURRENT_THD.Real_value            := INTERN.L1_CURRENT_THD;
	COM.HMI_OUTPUT_L1_CURRENT_THD.Real_value              := INTERN.L1_CURRENT_THD;
	COM.WEBVISU_OUTPUT_L1_CURRENT_THD.Real_value              := INTERN.L1_CURRENT_THD;
	COM.SCADA_OUTPUT_L1_MAX_LOAD.Real_value               := INTERN.L1_MAX_LOAD;
	COM.HMI_OUTPUT_L1_MAX_LOAD.Real_value                 := INTERN.L1_MAX_LOAD;
	COM.WEBVISU_OUTPUT_L1_MAX_LOAD.Real_value                 := INTERN.L1_MAX_LOAD;
	COM.SCADA_OUTPUT_L1_L2_VOLTAGE_PHASE_ANGLE.Real_value := INTERN.L1_L2_VOLTAGE_PHASE_ANGLE;
	COM.HMI_OUTPUT_L1_L2_VOLTAGE_PHASE_ANGLE.Real_value   := INTERN.L1_L2_VOLTAGE_PHASE_ANGLE;
	COM.WEBVISU_OUTPUT_L1_L2_VOLTAGE_PHASE_ANGLE.Real_value   := INTERN.L1_L2_VOLTAGE_PHASE_ANGLE;
	COM.SCADA_OUTPUT_L2_L3_VOLTAGE.Real_value             := INTERN.L2_L3_VOLTAGE;
	COM.HMI_OUTPUT_L2_L3_VOLTAGE.Real_value               := INTERN.L2_L3_VOLTAGE;
	COM.WEBVISU_OUTPUT_L2_L3_VOLTAGE.Real_value               := INTERN.L2_L3_VOLTAGE;
	COM.SCADA_OUTPUT_L2_N_VOLTAGE.Real_value              := INTERN.L2_N_VOLTAGE;
	COM.HMI_OUTPUT_L2_N_VOLTAGE.Real_value                := INTERN.L2_N_VOLTAGE;
	COM.WEBVISU_OUTPUT_L2_N_VOLTAGE.Real_value                := INTERN.L2_N_VOLTAGE;
	COM.SCADA_OUTPUT_L2_CURRENT.Real_value                := INTERN.L2_CURRENT;
	COM.HMI_OUTPUT_L2_CURRENT.Real_value                  := INTERN.L2_CURRENT;
	COM.WEBVISU_OUTPUT_L2_CURRENT.Real_value                  := INTERN.L2_CURRENT;
	COM.SCADA_OUTPUT_L2_ACTIVE_POWER.Real_value           := INTERN.L2_ACTIVE_POWER;
	COM.HMI_OUTPUT_L2_ACTIVE_POWER.Real_value             := INTERN.L2_ACTIVE_POWER;
	COM.WEBVISU_OUTPUT_L2_ACTIVE_POWER.Real_value             := INTERN.L2_ACTIVE_POWER;
	COM.SCADA_OUTPUT_L2_APPARENT_POWER.Real_value         := INTERN.L2_APPARENT_POWER;
	COM.HMI_OUTPUT_L2_APPARENT_POWER.Real_value           := INTERN.L2_APPARENT_POWER;
	COM.WEBVISU_OUTPUT_L2_APPARENT_POWER.Real_value           := INTERN.L2_APPARENT_POWER;
	COM.SCADA_OUTPUT_L2_REACTIVE_POWER.Real_value         := INTERN.L2_REACTIVE_POWER;
	COM.HMI_OUTPUT_L2_REACTIVE_POWER.Real_value           := INTERN.L2_REACTIVE_POWER;
	COM.WEBVISU_OUTPUT_L2_REACTIVE_POWER.Real_value           := INTERN.L2_REACTIVE_POWER;
	COM.SCADA_OUTPUT_L2_CURRENT_PHASE_ANGLE.Real_value    := INTERN.L2_CURRENT_PHASE_ANGLE;
	COM.HMI_OUTPUT_L2_CURRENT_PHASE_ANGLE.Real_value      := INTERN.L2_CURRENT_PHASE_ANGLE;
	COM.WEBVISU_OUTPUT_L2_CURRENT_PHASE_ANGLE.Real_value      := INTERN.L2_CURRENT_PHASE_ANGLE;
	COM.SCADA_OUTPUT_L2_POWER_FACTOR.Real_value           := INTERN.L2_POWER_FACTOR;
	COM.HMI_OUTPUT_L2_POWER_FACTOR.Real_value             := INTERN.L2_POWER_FACTOR;
	COM.WEBVISU_OUTPUT_L2_POWER_FACTOR.Real_value             := INTERN.L2_POWER_FACTOR;
	COM.SCADA_OUTPUT_L2_VOLTAGE_THD.Real_value            := INTERN.L2_VOLTAGE_THD;
	COM.HMI_OUTPUT_L2_VOLTAGE_THD.Real_value              := INTERN.L2_VOLTAGE_THD;
	COM.WEBVISU_OUTPUT_L2_VOLTAGE_THD.Real_value              := INTERN.L2_VOLTAGE_THD;
	COM.SCADA_OUTPUT_L2_CURRENT_THD.Real_value            := INTERN.L2_CURRENT_THD;
	COM.HMI_OUTPUT_L2_CURRENT_THD.Real_value              := INTERN.L2_CURRENT_THD;
	COM.WEBVISU_OUTPUT_L2_CURRENT_THD.Real_value              := INTERN.L2_CURRENT_THD;
	COM.SCADA_OUTPUT_L2_MAX_LOAD.Real_value               := INTERN.L2_MAX_LOAD;
	COM.HMI_OUTPUT_L2_MAX_LOAD.Real_value                 := INTERN.L2_MAX_LOAD;
	COM.WEBVISU_OUTPUT_L2_MAX_LOAD.Real_value                 := INTERN.L2_MAX_LOAD;
	COM.SCADA_OUTPUT_L1_L3_VOLTAGE_PHASE_ANGLE.Real_value := INTERN.L1_L3_VOLTAGE_PHASE_ANGLE;
	COM.HMI_OUTPUT_L1_L3_VOLTAGE_PHASE_ANGLE.Real_value   := INTERN.L1_L3_VOLTAGE_PHASE_ANGLE;
	COM.WEBVISU_OUTPUT_L1_L3_VOLTAGE_PHASE_ANGLE.Real_value   := INTERN.L1_L3_VOLTAGE_PHASE_ANGLE;
	COM.SCADA_OUTPUT_L3_L1_VOLTAGE.Real_value             := INTERN.L3_L1_VOLTAGE;
	COM.HMI_OUTPUT_L3_L1_VOLTAGE.Real_value               := INTERN.L3_L1_VOLTAGE;
	COM.WEBVISU_OUTPUT_L3_L1_VOLTAGE.Real_value               := INTERN.L3_L1_VOLTAGE;
	COM.SCADA_OUTPUT_L3_N_VOLTAGE.Real_value              := INTERN.L3_N_VOLTAGE;
	COM.HMI_OUTPUT_L3_N_VOLTAGE.Real_value                := INTERN.L3_N_VOLTAGE;
	COM.WEBVISU_OUTPUT_L3_N_VOLTAGE.Real_value                := INTERN.L3_N_VOLTAGE;
	COM.SCADA_OUTPUT_L3_CURRENT.Real_value                := INTERN.L3_CURRENT;
	COM.HMI_OUTPUT_L3_CURRENT.Real_value                  := INTERN.L3_CURRENT;
	COM.WEBVISU_OUTPUT_L3_CURRENT.Real_value                  := INTERN.L3_CURRENT;
	COM.SCADA_OUTPUT_L3_ACTIVE_POWER.Real_value           := INTERN.L3_ACTIVE_POWER;
	COM.HMI_OUTPUT_L3_ACTIVE_POWER.Real_value             := INTERN.L3_ACTIVE_POWER;
	COM.WEBVISU_OUTPUT_L3_ACTIVE_POWER.Real_value             := INTERN.L3_ACTIVE_POWER;
	COM.SCADA_OUTPUT_L3_APPARENT_POWER.Real_value         := INTERN.L3_APPARENT_POWER;
	COM.HMI_OUTPUT_L3_APPARENT_POWER.Real_value           := INTERN.L3_APPARENT_POWER;
	COM.WEBVISU_OUTPUT_L3_APPARENT_POWER.Real_value           := INTERN.L3_APPARENT_POWER;
	COM.SCADA_OUTPUT_L3_REACTIVE_POWER.Real_value         := INTERN.L3_REACTIVE_POWER;
	COM.HMI_OUTPUT_L3_REACTIVE_POWER.Real_value           := INTERN.L3_REACTIVE_POWER;
	COM.WEBVISU_OUTPUT_L3_REACTIVE_POWER.Real_value           := INTERN.L3_REACTIVE_POWER;
	COM.SCADA_OUTPUT_L3_CURRENT_PHASE_ANGLE.Real_value    := INTERN.L3_CURRENT_PHASE_ANGLE;
	COM.HMI_OUTPUT_L3_CURRENT_PHASE_ANGLE.Real_value      := INTERN.L3_CURRENT_PHASE_ANGLE;
	COM.WEBVISU_OUTPUT_L3_CURRENT_PHASE_ANGLE.Real_value      := INTERN.L3_CURRENT_PHASE_ANGLE;
	COM.SCADA_OUTPUT_L3_POWER_FACTOR.Real_value           := INTERN.L3_POWER_FACTOR;
	COM.HMI_OUTPUT_L3_POWER_FACTOR.Real_value             := INTERN.L3_POWER_FACTOR;
	COM.WEBVISU_OUTPUT_L3_POWER_FACTOR.Real_value             := INTERN.L3_POWER_FACTOR;
	COM.SCADA_OUTPUT_L3_VOLTAGE_THD.Real_value            := INTERN.L3_VOLTAGE_THD;
	COM.HMI_OUTPUT_L3_VOLTAGE_THD.Real_value              := INTERN.L3_VOLTAGE_THD;
	COM.WEBVISU_OUTPUT_L3_VOLTAGE_THD.Real_value              := INTERN.L3_VOLTAGE_THD;
	COM.SCADA_OUTPUT_L3_CURRENT_THD.Real_value            := INTERN.L3_CURRENT_THD;
	COM.HMI_OUTPUT_L3_CURRENT_THD.Real_value              := INTERN.L3_CURRENT_THD;
	COM.WEBVISU_OUTPUT_L3_CURRENT_THD.Real_value              := INTERN.L3_CURRENT_THD;
	COM.SCADA_OUTPUT_L3_MAX_LOAD.Real_value               := INTERN.L3_MAX_LOAD;
	COM.HMI_OUTPUT_L3_MAX_LOAD.Real_value                 := INTERN.L3_MAX_LOAD;
	COM.WEBVISU_OUTPUT_L3_MAX_LOAD.Real_value                 := INTERN.L3_MAX_LOAD;
	COM.SCADA_OUTPUT_INTERNAL_TEMPERATURE.Real_value      := INTERN.INTERNAL_TEMPERATURE;
	COM.HMI_OUTPUT_INTERNAL_TEMPERATURE.Real_value        := INTERN.INTERNAL_TEMPERATURE;
	COM.WEBVISU_OUTPUT_INTERNAL_TEMPERATURE.Real_value        := INTERN.INTERNAL_TEMPERATURE;
	COM.SCADA_OUTPUT_ACTIVE_ENERGY.Real_value             := INTERN.ACTIVE_ENERGY;
	COM.HMI_OUTPUT_ACTIVE_ENERGY.Real_value               := INTERN.ACTIVE_ENERGY;
	COM.WEBVISU_OUTPUT_ACTIVE_ENERGY.Real_value               := INTERN.ACTIVE_ENERGY;
	COM.SCADA_OUTPUT_APPARENT_ENERGY.Real_value           := INTERN.APPARENT_ENERGY;
	COM.HMI_OUTPUT_APPARENT_ENERGY.Real_value             := INTERN.APPARENT_ENERGY;
	COM.WEBVISU_OUTPUT_APPARENT_ENERGY.Real_value             := INTERN.APPARENT_ENERGY;
	COM.SCADA_OUTPUT_REACTIVE_ENERGY.Real_value           := INTERN.REACTIVE_ENERGY;
	COM.HMI_OUTPUT_REACTIVE_ENERGY.Real_value             := INTERN.REACTIVE_ENERGY;
	COM.WEBVISU_OUTPUT_REACTIVE_ENERGY.Real_value             := INTERN.REACTIVE_ENERGY;
	COM.SCADA_OUTPUT_TOTAL_ACTIVE_POWER.Real_value        := INTERN.TOTAL_ACTIVE_POWER;
	COM.HMI_OUTPUT_TOTAL_ACTIVE_POWER.Real_value          := INTERN.TOTAL_ACTIVE_POWER;
	COM.WEBVISU_OUTPUT_TOTAL_ACTIVE_POWER.Real_value          := INTERN.TOTAL_ACTIVE_POWER;
	COM.SCADA_OUTPUT_TOTAL_APPARENT_POWER.Real_value      := INTERN.TOTAL_APPARENT_POWER;
	COM.HMI_OUTPUT_TOTAL_APPARENT_POWER.Real_value        := INTERN.TOTAL_APPARENT_POWER;
	COM.WEBVISU_OUTPUT_TOTAL_APPARENT_POWER.Real_value        := INTERN.TOTAL_APPARENT_POWER;
	COM.SCADA_OUTPUT_TOTAL_REACTIVE_POWER.Real_value      := INTERN.TOTAL_REACTIVE_POWER;
	COM.HMI_OUTPUT_TOTAL_REACTIVE_POWER.Real_value        := INTERN.TOTAL_REACTIVE_POWER;
	COM.WEBVISU_OUTPUT_TOTAL_REACTIVE_POWER.Real_value        := INTERN.TOTAL_REACTIVE_POWER;
	COM.SCADA_OUTPUT_ALL_PHASE_POWER_FACTOR.Real_value    := INTERN.ALL_PHASE_POWER_FACTOR;
	COM.HMI_OUTPUT_ALL_PHASE_POWER_FACTOR.Real_value      := INTERN.ALL_PHASE_POWER_FACTOR;
	COM.WEBVISU_OUTPUT_ALL_PHASE_POWER_FACTOR.Real_value      := INTERN.ALL_PHASE_POWER_FACTOR;


          
END_FUNCTION_BLOCK

FUNCTION_BLOCK FB_INST_DIP1500
  VAR_IN_OUT
    PA : DUT_PA_DIP1500;  (* Parameters (persistent, GVL_PA) *)
    COM : DUT_COM_DIP1500;  (* Communication : Modbus RTU (COM_), SCADA FUXA (SCADA_), HMI (HMI_) *)
    EXC : DUT_EXC_DIP1500;  (* Exchanges : other equipment (EXC_), functional units (UPI_) *)
    IO : DUT_IO_DIP1500;  (* Wired PLC I/O *)
  END_VAR
  VAR
    INTERN : DUT_INT_DIP1500;  (* Internal variables *)
    TON_PULSE : TON;  (* Square wave timer *)
    TOF_CMD_WINDOW : TOF;  (* Command write window *)
    R_TRIG_FLASH : R_TRIG;  (* Flash save request edge *)
    TP_FLASH : TP;  (* Flash save pulse *)
  END_VAR

            
//==============================================================================
// FB_INST_DIP1500
// Kamoer DIP1500 peristaltic pump, Modbus RTU, 32-bit low word first (CDAB)
// 1. INPUTS     : requests, control mode, command source, equipment feedback -> INTERN
// 2. PROCESSING : on INTERN only
// 3. OUTPUTS    : INTERN -> COM / IO / EXC
// Parameters    : pump configuration in PA (persistent), changed from the active local supervision
// Control mode  : local WEBVISU > local HMI > local FUXA > auto (functional units)
//==============================================================================

//------------------------------------------------------------------------------
// 1. INPUTS
//------------------------------------------------------------------------------
	//--- Control mode requests (WEBVISU, HMI, FUXA, global UPI)
	INTERN.FUXA_LOCAL_REQUEST := COM.SCADA_INPUT_LOCAL_REQUEST;
	INTERN.FUXA_AUTO_REQUEST  := COM.SCADA_INPUT_AUTO_REQUEST;
	INTERN.HMI_LOCAL_REQUEST  := COM.HMI_INPUT_LOCAL_REQUEST;
	INTERN.HMI_AUTO_REQUEST   := COM.HMI_INPUT_AUTO_REQUEST;
	INTERN.GLOBAL_LOCAL_FUXA  := EXC.UPI_INPUT_GLOBAL_LOCAL_FUXA;
	INTERN.GLOBAL_LOCAL_HMI   := EXC.UPI_INPUT_GLOBAL_LOCAL_HMI;
	INTERN.WEBVISU_LOCAL_REQUEST := COM.WEBVISU_INPUT_LOCAL_REQUEST;
	INTERN.WEBVISU_AUTO_REQUEST  := COM.WEBVISU_INPUT_AUTO_REQUEST;
	INTERN.GLOBAL_LOCAL_WEBVISU  := EXC.UPI_INPUT_GLOBAL_LOCAL_WEBVISU;

	//--- Control mode
	// Individual memories : set by the local request, reset by the auto request (auto wins if both)
	IF INTERN.WEBVISU_LOCAL_REQUEST THEN
		INTERN.LOCAL_WEBVISU_INDIVIDUAL := TRUE;
	END_IF
	IF INTERN.WEBVISU_AUTO_REQUEST THEN
		INTERN.LOCAL_WEBVISU_INDIVIDUAL := FALSE;
	END_IF
	IF INTERN.HMI_LOCAL_REQUEST THEN
		INTERN.LOCAL_HMI_INDIVIDUAL := TRUE;
	END_IF
	IF INTERN.HMI_AUTO_REQUEST THEN
		INTERN.LOCAL_HMI_INDIVIDUAL := FALSE;
	END_IF
	IF INTERN.FUXA_LOCAL_REQUEST THEN
		INTERN.LOCAL_FUXA_INDIVIDUAL := TRUE;
	END_IF
	IF INTERN.FUXA_AUTO_REQUEST THEN
		INTERN.LOCAL_FUXA_INDIVIDUAL := FALSE;
	END_IF

	// Resulting mode : individual OR global, WEBVISU > HMI > FUXA > auto
	INTERN.LOCAL_WEBVISU := INTERN.LOCAL_WEBVISU_INDIVIDUAL OR INTERN.GLOBAL_LOCAL_WEBVISU;
	INTERN.LOCAL_HMI     := (INTERN.LOCAL_HMI_INDIVIDUAL OR INTERN.GLOBAL_LOCAL_HMI) AND NOT INTERN.LOCAL_WEBVISU;
	INTERN.LOCAL_FUXA    := (INTERN.LOCAL_FUXA_INDIVIDUAL OR INTERN.GLOBAL_LOCAL_FUXA) AND NOT INTERN.LOCAL_WEBVISU AND NOT INTERN.LOCAL_HMI;
	INTERN.AUTO          := NOT INTERN.LOCAL_WEBVISU AND NOT INTERN.LOCAL_HMI AND NOT INTERN.LOCAL_FUXA;

	//--- Command source : local WEBVISU > local HMI > local FUXA > auto (UPI)
	IF INTERN.LOCAL_WEBVISU THEN
		INTERN.CMD_RUN            := COM.WEBVISU_INPUT_MOTOR_START_STOP;
		INTERN.CMD_CLOCKWISE      := COM.WEBVISU_INPUT_MOTOR_DIRECTION;
		INTERN.CMD_VOLUME_MODE    := COM.WEBVISU_INPUT_OPERATION_MODE;
		INTERN.CMD_SPEED          := COM.WEBVISU_INPUT_MOTOR_SPEED.Real_value;
		INTERN.CMD_RUN_SETPOINT   := COM.WEBVISU_INPUT_RUN_TIME_OR_VOLUME_SETPOINT.Real_value;
		INTERN.PARAM_WRITE_ENABLE := COM.WEBVISU_INPUT_PARAM_WRITE_ENABLE;
		INTERN.FLASH_SAVE_REQUEST := COM.WEBVISU_INPUT_FLASH_SAVE;
	ELSIF INTERN.LOCAL_HMI THEN
		INTERN.CMD_RUN            := COM.HMI_INPUT_MOTOR_START_STOP;
		INTERN.CMD_CLOCKWISE      := COM.HMI_INPUT_MOTOR_DIRECTION;
		INTERN.CMD_VOLUME_MODE    := COM.HMI_INPUT_OPERATION_MODE;
		INTERN.CMD_SPEED          := COM.HMI_INPUT_MOTOR_SPEED.Real_value;
		INTERN.CMD_RUN_SETPOINT   := COM.HMI_INPUT_RUN_TIME_OR_VOLUME_SETPOINT.Real_value;
		INTERN.PARAM_WRITE_ENABLE := COM.HMI_INPUT_PARAM_WRITE_ENABLE;
		INTERN.FLASH_SAVE_REQUEST := COM.HMI_INPUT_FLASH_SAVE;
	ELSIF INTERN.LOCAL_FUXA THEN
		INTERN.CMD_RUN            := COM.SCADA_INPUT_MOTOR_START_STOP;
		INTERN.CMD_CLOCKWISE      := COM.SCADA_INPUT_MOTOR_DIRECTION;
		INTERN.CMD_VOLUME_MODE    := COM.SCADA_INPUT_OPERATION_MODE;
		INTERN.CMD_SPEED          := COM.SCADA_INPUT_MOTOR_SPEED.Real_value;
		INTERN.CMD_RUN_SETPOINT   := COM.SCADA_INPUT_RUN_TIME_OR_VOLUME_SETPOINT.Real_value;
		INTERN.PARAM_WRITE_ENABLE := COM.SCADA_INPUT_PARAM_WRITE_ENABLE;
		INTERN.FLASH_SAVE_REQUEST := COM.SCADA_INPUT_FLASH_SAVE;
	ELSE
		// Auto : functional units (UPI)
		INTERN.CMD_RUN            := EXC.UPI_INPUT_RUN;
		INTERN.CMD_CLOCKWISE      := EXC.UPI_INPUT_CLOCKWISE;
		INTERN.CMD_VOLUME_MODE    := EXC.UPI_INPUT_VOLUME_MODE;
		INTERN.CMD_SPEED          := EXC.UPI_INPUT_SPEED;
		INTERN.CMD_RUN_SETPOINT   := EXC.UPI_INPUT_RUN_SETPOINT;
		INTERN.PARAM_WRITE_ENABLE := FALSE;                        // configuration is never written in auto
		INTERN.FLASH_SAVE_REQUEST := FALSE;
	END_IF

	//--- Parameter source : values typed in the active local supervision (nothing in auto)
	IF INTERN.LOCAL_WEBVISU THEN
		INTERN.SRC_MAX_MOTOR_SPEED         := COM.WEBVISU_INPUT_MAX_MOTOR_SPEED.Real_value;
		INTERN.SRC_CALIBRATION_COEFFICIENT := COM.WEBVISU_INPUT_FLOW_RATE_OR_SPEED_CALIBRATION_COEFFICIENT.Real_value;
		INTERN.SRC_FOOT_SWITCH_INPUT_MODE  := COM.WEBVISU_INPUT_FOOT_SWITCH_INPUT_MODE;
		INTERN.SRC_LIQUID_LEVEL_INPUT_MODE := COM.WEBVISU_INPUT_LIQUID_LEVEL_INPUT_MODE;
		INTERN.SRC_STATE_OUTPUT_MODE       := COM.WEBVISU_INPUT_STATE_OUTPUT_MODE;
		INTERN.SRC_COMMUNICATION_ADDRESS   := COM.WEBVISU_INPUT_COMMUNICATION_ADDRESS;
		INTERN.SRC_BAUD_RATE_INDEX         := COM.WEBVISU_INPUT_BAUD_RATE_INDEX;
	ELSIF INTERN.LOCAL_HMI THEN
		INTERN.SRC_MAX_MOTOR_SPEED         := COM.HMI_INPUT_MAX_MOTOR_SPEED.Real_value;
		INTERN.SRC_CALIBRATION_COEFFICIENT := COM.HMI_INPUT_FLOW_RATE_OR_SPEED_CALIBRATION_COEFFICIENT.Real_value;
		INTERN.SRC_FOOT_SWITCH_INPUT_MODE  := COM.HMI_INPUT_FOOT_SWITCH_INPUT_MODE;
		INTERN.SRC_LIQUID_LEVEL_INPUT_MODE := COM.HMI_INPUT_LIQUID_LEVEL_INPUT_MODE;
		INTERN.SRC_STATE_OUTPUT_MODE       := COM.HMI_INPUT_STATE_OUTPUT_MODE;
		INTERN.SRC_COMMUNICATION_ADDRESS   := COM.HMI_INPUT_COMMUNICATION_ADDRESS;
		INTERN.SRC_BAUD_RATE_INDEX         := COM.HMI_INPUT_BAUD_RATE_INDEX;
	ELSIF INTERN.LOCAL_FUXA THEN
		INTERN.SRC_MAX_MOTOR_SPEED         := COM.SCADA_INPUT_MAX_MOTOR_SPEED.Real_value;
		INTERN.SRC_CALIBRATION_COEFFICIENT := COM.SCADA_INPUT_FLOW_RATE_OR_SPEED_CALIBRATION_COEFFICIENT.Real_value;
		INTERN.SRC_FOOT_SWITCH_INPUT_MODE  := COM.SCADA_INPUT_FOOT_SWITCH_INPUT_MODE;
		INTERN.SRC_LIQUID_LEVEL_INPUT_MODE := COM.SCADA_INPUT_LIQUID_LEVEL_INPUT_MODE;
		INTERN.SRC_STATE_OUTPUT_MODE       := COM.SCADA_INPUT_STATE_OUTPUT_MODE;
		INTERN.SRC_COMMUNICATION_ADDRESS   := COM.SCADA_INPUT_COMMUNICATION_ADDRESS;
		INTERN.SRC_BAUD_RATE_INDEX         := COM.SCADA_INPUT_BAUD_RATE_INDEX;
	END_IF

	//--- COM : input registers 0x3001..0x3005
	INTERN.FBK_FIRMWARE_VERSION := COM.COM_INPUT_IR[0];
	INTERN.FBK_HARDWARE_VERSION := COM.COM_INPUT_IR[1];
	INTERN.FBK_TEMPERATURE      := COM.COM_INPUT_IR[2];
	INTERN.FBK_LEVEL_ALARM      := COM.COM_INPUT_IR[3];
	INTERN.FBK_DIGITAL_OUTPUT   := COM.COM_INPUT_IR[4];

	//--- COM : run counters 0x4007..0x400A (format depends on mode)
	IF INTERN.CMD_VOLUME_MODE THEN
		// Volume mode : 32-bit REAL (ml)
		INTERN.FBK_RUN_ACTUAL := FNC_WORDS_TO_REAL(High_word := COM.COM_INPUT_HR_COUNTERS[1], Low_word := COM.COM_INPUT_HR_COUNTERS[0]);
		INTERN.FBK_RUN_TOTAL  := FNC_WORDS_TO_REAL(High_word := COM.COM_INPUT_HR_COUNTERS[3], Low_word := COM.COM_INPUT_HR_COUNTERS[2]);
	ELSE
		// Time mode : 32-bit UDINT (ms)
		INTERN.UDINT_TEMP     := SHL(WORD_TO_UDINT(COM.COM_INPUT_HR_COUNTERS[1]), 16) OR WORD_TO_UDINT(COM.COM_INPUT_HR_COUNTERS[0]);
		INTERN.FBK_RUN_ACTUAL := UDINT_TO_REAL(INTERN.UDINT_TEMP);
		INTERN.UDINT_TEMP     := SHL(WORD_TO_UDINT(COM.COM_INPUT_HR_COUNTERS[3]), 16) OR WORD_TO_UDINT(COM.COM_INPUT_HR_COUNTERS[2]);
		INTERN.FBK_RUN_TOTAL  := UDINT_TO_REAL(INTERN.UDINT_TEMP);
	END_IF


//------------------------------------------------------------------------------
// 2. PROCESSING
//------------------------------------------------------------------------------
	//--- Parameters (PA) : a value changed in the active supervision is saved in PA
	// PA is persistent : it keeps its value after a restart or a download. Default = declaration value.
	// The cycle where the source changes is ignored, so switching mode never overwrites PA.
	INTERN.SOURCE_CHANGED := (INTERN.LOCAL_WEBVISU <> INTERN.PREV_LOCAL_WEBVISU)
	                         OR (INTERN.LOCAL_HMI <> INTERN.PREV_LOCAL_HMI)
	                         OR (INTERN.LOCAL_FUXA <> INTERN.PREV_LOCAL_FUXA);
	INTERN.PREV_LOCAL_WEBVISU := INTERN.LOCAL_WEBVISU;
	INTERN.PREV_LOCAL_HMI     := INTERN.LOCAL_HMI;
	INTERN.PREV_LOCAL_FUXA    := INTERN.LOCAL_FUXA;

	IF NOT INTERN.SOURCE_CHANGED THEN
		IF INTERN.SRC_MAX_MOTOR_SPEED <> INTERN.PREV_SRC_MAX_MOTOR_SPEED THEN
			PA.MAX_MOTOR_SPEED := INTERN.SRC_MAX_MOTOR_SPEED;
		END_IF
		IF INTERN.SRC_CALIBRATION_COEFFICIENT <> INTERN.PREV_SRC_CALIBRATION_COEFFICIENT THEN
			PA.CALIBRATION_COEFFICIENT := INTERN.SRC_CALIBRATION_COEFFICIENT;
		END_IF
		IF INTERN.SRC_FOOT_SWITCH_INPUT_MODE <> INTERN.PREV_SRC_FOOT_SWITCH_INPUT_MODE THEN
			PA.FOOT_SWITCH_INPUT_MODE := INTERN.SRC_FOOT_SWITCH_INPUT_MODE;
		END_IF
		IF INTERN.SRC_LIQUID_LEVEL_INPUT_MODE <> INTERN.PREV_SRC_LIQUID_LEVEL_INPUT_MODE THEN
			PA.LIQUID_LEVEL_INPUT_MODE := INTERN.SRC_LIQUID_LEVEL_INPUT_MODE;
		END_IF
		IF INTERN.SRC_STATE_OUTPUT_MODE <> INTERN.PREV_SRC_STATE_OUTPUT_MODE THEN
			PA.STATE_OUTPUT_MODE := INTERN.SRC_STATE_OUTPUT_MODE;
		END_IF
		IF INTERN.SRC_COMMUNICATION_ADDRESS <> INTERN.PREV_SRC_COMMUNICATION_ADDRESS THEN
			PA.COMMUNICATION_ADDRESS := INTERN.SRC_COMMUNICATION_ADDRESS;
		END_IF
		IF INTERN.SRC_BAUD_RATE_INDEX <> INTERN.PREV_SRC_BAUD_RATE_INDEX THEN
			PA.BAUD_RATE_INDEX := INTERN.SRC_BAUD_RATE_INDEX;
		END_IF
	END_IF

	INTERN.PREV_SRC_MAX_MOTOR_SPEED         := INTERN.SRC_MAX_MOTOR_SPEED;
	INTERN.PREV_SRC_CALIBRATION_COEFFICIENT := INTERN.SRC_CALIBRATION_COEFFICIENT;
	INTERN.PREV_SRC_FOOT_SWITCH_INPUT_MODE  := INTERN.SRC_FOOT_SWITCH_INPUT_MODE;
	INTERN.PREV_SRC_LIQUID_LEVEL_INPUT_MODE := INTERN.SRC_LIQUID_LEVEL_INPUT_MODE;
	INTERN.PREV_SRC_STATE_OUTPUT_MODE       := INTERN.SRC_STATE_OUTPUT_MODE;
	INTERN.PREV_SRC_COMMUNICATION_ADDRESS   := INTERN.SRC_COMMUNICATION_ADDRESS;
	INTERN.PREV_SRC_BAUD_RATE_INDEX         := INTERN.SRC_BAUD_RATE_INDEX;

	//--- Parameters used by the pump : always from PA
	INTERN.CMD_MAX_SPEED      := PA.MAX_MOTOR_SPEED;
	INTERN.CMD_CALIB_COEF     := PA.CALIBRATION_COEFFICIENT;
	INTERN.CMD_FOOT_MODE      := PA.FOOT_SWITCH_INPUT_MODE;
	INTERN.CMD_LEVEL_MODE     := PA.LIQUID_LEVEL_INPUT_MODE;
	INTERN.CMD_STATE_OUT_MODE := PA.STATE_OUTPUT_MODE;
	INTERN.CMD_ADDRESS        := PA.COMMUNICATION_ADDRESS;
	INTERN.CMD_BAUD_INDEX     := PA.BAUD_RATE_INDEX;

	//--- Parameter validity
	INTERN.PARAM_VALID := (WORD_TO_UINT(INTERN.CMD_ADDRESS) >= 1) AND (WORD_TO_UINT(INTERN.CMD_ADDRESS) <= 31)
	                      AND (WORD_TO_UINT(INTERN.CMD_BAUD_INDEX) <= 7)
	                      AND (INTERN.CMD_MAX_SPEED > 0.0) AND (INTERN.CMD_CALIB_COEF > 0.0);

	//--- Flash save : 1 s pulse on rising edge, only with valid parameters
	R_TRIG_FLASH(CLK := INTERN.FLASH_SAVE_REQUEST);
	TP_FLASH(IN := R_TRIG_FLASH.Q AND INTERN.PARAM_VALID, PT := T#1S);
	INTERN.CMD_SAVE_FLASH := TP_FLASH.Q;

	//--- Write triggers (rising edge channels)
	// Square wave 500 ms : each rising edge = one write request
	TON_PULSE(IN := NOT TON_PULSE.Q, PT := T#250MS);
	IF TON_PULSE.Q THEN
		INTERN.PULSE_500MS := NOT INTERN.PULSE_500MS;
	END_IF

	// Command trigger : automatic, 3 s of edges after any command change
	INTERN.CMD_CHANGED := (INTERN.CMD_RUN <> INTERN.PREV_RUN) OR (INTERN.CMD_CLOCKWISE <> INTERN.PREV_CLOCKWISE)
	                      OR (INTERN.CMD_VOLUME_MODE <> INTERN.PREV_VOLUME_MODE) OR (INTERN.CMD_SAVE_FLASH <> INTERN.PREV_SAVE_FLASH)
	                      OR (INTERN.CMD_SPEED <> INTERN.PREV_SPEED) OR (INTERN.CMD_MAX_SPEED <> INTERN.PREV_MAX_SPEED)
	                      OR (INTERN.CMD_RUN_SETPOINT <> INTERN.PREV_RUN_SETPOINT);
	INTERN.PREV_RUN          := INTERN.CMD_RUN;
	INTERN.PREV_CLOCKWISE    := INTERN.CMD_CLOCKWISE;
	INTERN.PREV_VOLUME_MODE  := INTERN.CMD_VOLUME_MODE;
	INTERN.PREV_SAVE_FLASH   := INTERN.CMD_SAVE_FLASH;
	INTERN.PREV_SPEED        := INTERN.CMD_SPEED;
	INTERN.PREV_MAX_SPEED    := INTERN.CMD_MAX_SPEED;
	INTERN.PREV_RUN_SETPOINT := INTERN.CMD_RUN_SETPOINT;

	TOF_CMD_WINDOW(IN := INTERN.CMD_CHANGED, PT := T#3S);
	INTERN.CMD_WINDOW  := TOF_CMD_WINDOW.Q;
	INTERN.CMD_TRIGGER := INTERN.CMD_WINDOW AND (INTERN.CMD_MAX_SPEED > 0.0) AND INTERN.PULSE_500MS;

	// Configuration trigger : only while writing is enabled and parameters are valid
	INTERN.CONFIG_TRIGGER := INTERN.PARAM_WRITE_ENABLE AND INTERN.PARAM_VALID AND INTERN.PULSE_500MS;


//------------------------------------------------------------------------------
// 3. OUTPUTS
//------------------------------------------------------------------------------
	//--- COM : control mode status to SCADA, HMI and WEBVISU
	COM.SCADA_OUTPUT_LOCAL_FUXA_ACTIVE := INTERN.LOCAL_FUXA;
	COM.SCADA_OUTPUT_LOCAL_HMI_ACTIVE  := INTERN.LOCAL_HMI;
	COM.HMI_OUTPUT_LOCAL_ACTIVE        := INTERN.LOCAL_HMI;
	COM.WEBVISU_OUTPUT_LOCAL_ACTIVE        := INTERN.LOCAL_WEBVISU;
	COM.WEBVISU_OUTPUT_LOCAL_HMI_ACTIVE  := INTERN.LOCAL_HMI;
	COM.WEBVISU_OUTPUT_LOCAL_FUXA_ACTIVE := INTERN.LOCAL_FUXA;

	//--- COM : Modbus RTU coils
	COM.COM_OUTPUT_COILS[0] := INTERN.CMD_RUN;           // 0x0001
	COM.COM_OUTPUT_COILS[1] := INTERN.CMD_CLOCKWISE;     // 0x0002
	COM.COM_OUTPUT_COILS[2] := INTERN.CMD_SAVE_FLASH;    // 0x0003
	COM.COM_OUTPUT_COILS[3] := INTERN.CMD_VOLUME_MODE;   // 0x0004

	//--- COM : Modbus RTU holding registers and write triggers
	// Command registers 0x4001..0x4006 (sent on the command trigger)
	FNC_REAL_TO_WORDS(Real_value := INTERN.CMD_SPEED,     High_word => COM.COM_OUTPUT_HR_CMD[1], Low_word => COM.COM_OUTPUT_HR_CMD[0]);   // 0x4001-4002
	FNC_REAL_TO_WORDS(Real_value := INTERN.CMD_MAX_SPEED, High_word => COM.COM_OUTPUT_HR_CMD[3], Low_word => COM.COM_OUTPUT_HR_CMD[2]);   // 0x4003-4004
	IF INTERN.CMD_VOLUME_MODE THEN
		// Run setpoint 0x4005-4006, volume mode : 32-bit REAL (ml)
		FNC_REAL_TO_WORDS(Real_value := INTERN.CMD_RUN_SETPOINT, High_word => COM.COM_OUTPUT_HR_CMD[5], Low_word => COM.COM_OUTPUT_HR_CMD[4]);
	ELSE
		// Run setpoint 0x4005-4006, time mode : 32-bit UDINT (ms)
		INTERN.UDINT_TEMP        := REAL_TO_UDINT(MAX(INTERN.CMD_RUN_SETPOINT, 0.0));
		COM.COM_OUTPUT_HR_CMD[4] := UDINT_TO_WORD(INTERN.UDINT_TEMP);
		COM.COM_OUTPUT_HR_CMD[5] := UDINT_TO_WORD(SHR(INTERN.UDINT_TEMP, 16));
	END_IF

	// Configuration registers 0x400B..0x4011 (sent on the configuration trigger), updated only while enabled and valid
	IF INTERN.PARAM_WRITE_ENABLE AND INTERN.PARAM_VALID THEN
		FNC_REAL_TO_WORDS(Real_value := INTERN.CMD_CALIB_COEF, High_word => COM.COM_OUTPUT_HR_CONFIG[1], Low_word => COM.COM_OUTPUT_HR_CONFIG[0]);   // 0x400B-400C
		COM.COM_OUTPUT_HR_CONFIG[2] := INTERN.CMD_FOOT_MODE;        // 0x400D
		COM.COM_OUTPUT_HR_CONFIG[3] := INTERN.CMD_LEVEL_MODE;       // 0x400E
		COM.COM_OUTPUT_HR_CONFIG[4] := INTERN.CMD_STATE_OUT_MODE;   // 0x400F
		COM.COM_OUTPUT_HR_CONFIG[5] := INTERN.CMD_ADDRESS;          // 0x4010
		COM.COM_OUTPUT_HR_CONFIG[6] := INTERN.CMD_BAUD_INDEX;       // 0x4011
	END_IF

	// Write triggers
	COM.COM_OUTPUT_CMD_TRIGGER    := INTERN.CMD_TRIGGER;
	COM.COM_OUTPUT_CONFIG_TRIGGER := INTERN.CONFIG_TRIGGER;

	//--- COM : feedback to SCADA, HMI and WEBVISU
	COM.SCADA_OUTPUT_FIRMWARE_VERSION                          := INTERN.FBK_FIRMWARE_VERSION;
	COM.HMI_OUTPUT_FIRMWARE_VERSION                            := INTERN.FBK_FIRMWARE_VERSION;
	COM.WEBVISU_OUTPUT_FIRMWARE_VERSION                            := INTERN.FBK_FIRMWARE_VERSION;
	COM.SCADA_OUTPUT_HARDWARE_VERSION                          := INTERN.FBK_HARDWARE_VERSION;
	COM.HMI_OUTPUT_HARDWARE_VERSION                            := INTERN.FBK_HARDWARE_VERSION;
	COM.WEBVISU_OUTPUT_HARDWARE_VERSION                            := INTERN.FBK_HARDWARE_VERSION;
	COM.SCADA_OUTPUT_TEMPERATURE                               := INTERN.FBK_TEMPERATURE;
	COM.HMI_OUTPUT_TEMPERATURE                                 := INTERN.FBK_TEMPERATURE;
	COM.WEBVISU_OUTPUT_TEMPERATURE                                 := INTERN.FBK_TEMPERATURE;
	COM.SCADA_OUTPUT_FLOAT_LEVEL_ALARM                         := INTERN.FBK_LEVEL_ALARM;
	COM.HMI_OUTPUT_FLOAT_LEVEL_ALARM                           := INTERN.FBK_LEVEL_ALARM;
	COM.WEBVISU_OUTPUT_FLOAT_LEVEL_ALARM                           := INTERN.FBK_LEVEL_ALARM;
	COM.SCADA_OUTPUT_DIGITAL_OUTPUT_VALUE                      := INTERN.FBK_DIGITAL_OUTPUT;
	COM.HMI_OUTPUT_DIGITAL_OUTPUT_VALUE                        := INTERN.FBK_DIGITAL_OUTPUT;
	COM.WEBVISU_OUTPUT_DIGITAL_OUTPUT_VALUE                        := INTERN.FBK_DIGITAL_OUTPUT;
	COM.SCADA_OUTPUT_REAL_TIME_RUN_TIME_OR_VOLUME.Real_value   := INTERN.FBK_RUN_ACTUAL;
	COM.HMI_OUTPUT_REAL_TIME_RUN_TIME_OR_VOLUME.Real_value     := INTERN.FBK_RUN_ACTUAL;
	COM.WEBVISU_OUTPUT_REAL_TIME_RUN_TIME_OR_VOLUME.Real_value     := INTERN.FBK_RUN_ACTUAL;
	COM.SCADA_OUTPUT_ACCUMULATED_RUN_TIME_OR_VOLUME.Real_value := INTERN.FBK_RUN_TOTAL;
	COM.HMI_OUTPUT_ACCUMULATED_RUN_TIME_OR_VOLUME.Real_value   := INTERN.FBK_RUN_TOTAL;
	COM.WEBVISU_OUTPUT_ACCUMULATED_RUN_TIME_OR_VOLUME.Real_value   := INTERN.FBK_RUN_TOTAL;


          
END_FUNCTION_BLOCK

FUNCTION_BLOCK FB_INST_DOSENSOR
  VAR_IN_OUT
    PA : DUT_PA_DOSENSOR;  (* Parameters (persistent, GVL_PA) *)
    COM : DUT_COM_DOSENSOR;  (* Communication : Modbus RTU (COM_), SCADA FUXA (SCADA_), HMI (HMI_) *)
    EXC : DUT_EXC_DOSENSOR;  (* Exchanges : other equipment (EXC_), functional units (UPI_) *)
    IO : DUT_IO_DOSENSOR;  (* Wired PLC I/O *)
  END_VAR
  VAR
    INTERN : DUT_INT_DOSENSOR;  (* Internal variables *)
    TP_CALIB_HIGH : TP;  (* High calibration pulse *)
    TP_CALIB_LOW : TP;  (* Low calibration pulse *)
    TP_CALIB_DONE : TP;  (* Calibration done message *)
  END_VAR

            
//==============================================================================
// FB_INST_DOSENSOR
// Dissolved oxygen sensor, analog signal + fault input + 2 calibration outputs
// 1. INPUTS     : requests, control mode, command source, equipment feedback -> INTERN
// 2. PROCESSING : on INTERN only
// 3. OUTPUTS    : INTERN -> COM / IO / EXC
// Control mode  : local WEBVISU > local HMI > local FUXA > auto (functional units)
//==============================================================================

//------------------------------------------------------------------------------
// 1. INPUTS
//------------------------------------------------------------------------------
	//--- Control mode requests (WEBVISU, HMI, FUXA, global UPI)
	INTERN.FUXA_LOCAL_REQUEST := COM.SCADA_INPUT_LOCAL_REQUEST;
	INTERN.FUXA_AUTO_REQUEST  := COM.SCADA_INPUT_AUTO_REQUEST;
	INTERN.HMI_LOCAL_REQUEST  := COM.HMI_INPUT_LOCAL_REQUEST;
	INTERN.HMI_AUTO_REQUEST   := COM.HMI_INPUT_AUTO_REQUEST;
	INTERN.GLOBAL_LOCAL_FUXA  := EXC.UPI_INPUT_GLOBAL_LOCAL_FUXA;
	INTERN.GLOBAL_LOCAL_HMI   := EXC.UPI_INPUT_GLOBAL_LOCAL_HMI;
	INTERN.WEBVISU_LOCAL_REQUEST := COM.WEBVISU_INPUT_LOCAL_REQUEST;
	INTERN.WEBVISU_AUTO_REQUEST  := COM.WEBVISU_INPUT_AUTO_REQUEST;
	INTERN.GLOBAL_LOCAL_WEBVISU  := EXC.UPI_INPUT_GLOBAL_LOCAL_WEBVISU;
	//--- Control mode
	// Individual memories : set by the local request, reset by the auto request (auto wins if both)
	IF INTERN.WEBVISU_LOCAL_REQUEST THEN
		INTERN.LOCAL_WEBVISU_INDIVIDUAL := TRUE;
	END_IF
	IF INTERN.WEBVISU_AUTO_REQUEST THEN
		INTERN.LOCAL_WEBVISU_INDIVIDUAL := FALSE;
	END_IF
	IF INTERN.HMI_LOCAL_REQUEST THEN
		INTERN.LOCAL_HMI_INDIVIDUAL := TRUE;
	END_IF
	IF INTERN.HMI_AUTO_REQUEST THEN
		INTERN.LOCAL_HMI_INDIVIDUAL := FALSE;
	END_IF
	IF INTERN.FUXA_LOCAL_REQUEST THEN
		INTERN.LOCAL_FUXA_INDIVIDUAL := TRUE;
	END_IF
	IF INTERN.FUXA_AUTO_REQUEST THEN
		INTERN.LOCAL_FUXA_INDIVIDUAL := FALSE;
	END_IF

	// Resulting mode : individual OR global, WEBVISU > HMI > FUXA > auto
	INTERN.LOCAL_WEBVISU := INTERN.LOCAL_WEBVISU_INDIVIDUAL OR INTERN.GLOBAL_LOCAL_WEBVISU;
	INTERN.LOCAL_HMI     := (INTERN.LOCAL_HMI_INDIVIDUAL OR INTERN.GLOBAL_LOCAL_HMI) AND NOT INTERN.LOCAL_WEBVISU;
	INTERN.LOCAL_FUXA    := (INTERN.LOCAL_FUXA_INDIVIDUAL OR INTERN.GLOBAL_LOCAL_FUXA) AND NOT INTERN.LOCAL_WEBVISU AND NOT INTERN.LOCAL_HMI;
	INTERN.AUTO          := NOT INTERN.LOCAL_WEBVISU AND NOT INTERN.LOCAL_HMI AND NOT INTERN.LOCAL_FUXA;

	//--- Command source : calibration requests
	IF INTERN.LOCAL_WEBVISU THEN
		INTERN.CALIB_HIGH_REQUEST := COM.WEBVISU_INPUT_CALIBRATION_HIGH;
		INTERN.CALIB_LOW_REQUEST  := COM.WEBVISU_INPUT_CALIBRATION_LOW;
	ELSIF INTERN.LOCAL_HMI THEN
		INTERN.CALIB_HIGH_REQUEST := COM.HMI_INPUT_CALIBRATION_HIGH;
		INTERN.CALIB_LOW_REQUEST  := COM.HMI_INPUT_CALIBRATION_LOW;
	ELSIF INTERN.LOCAL_FUXA THEN
		INTERN.CALIB_HIGH_REQUEST := COM.SCADA_INPUT_CALIBRATION_HIGH;
		INTERN.CALIB_LOW_REQUEST  := COM.SCADA_INPUT_CALIBRATION_LOW;
	ELSE
		// Auto : functional units (UPI)
		INTERN.CALIB_HIGH_REQUEST := FALSE;
		INTERN.CALIB_LOW_REQUEST  := FALSE;
	END_IF

	//--- IO
	INTERN.SIGNAL_RAW := IO.INPUT_SIGNAL;
	INTERN.FAULT      := IO.INPUT_SENSOR_FAULT;


//------------------------------------------------------------------------------
// 2. PROCESSING
//------------------------------------------------------------------------------
	//--- Signal scaling
	INTERN.SIGNAL := (DWORD_TO_REAL(INTERN.SIGNAL_RAW * 40) / 65535) - 8;

	//--- Calibration : 1 s pulse to the sensor, 5 s "done" message
	TP_CALIB_HIGH(IN := INTERN.CALIB_HIGH_REQUEST, PT := T#1S);
	TP_CALIB_LOW(IN := INTERN.CALIB_LOW_REQUEST, PT := T#1S);
	TP_CALIB_DONE(IN := TP_CALIB_HIGH.Q OR TP_CALIB_LOW.Q, PT := T#5S);

	INTERN.CALIB_HIGH := TP_CALIB_HIGH.Q;
	INTERN.CALIB_LOW  := TP_CALIB_LOW.Q;
	INTERN.CALIB_DONE := TP_CALIB_DONE.Q;


//------------------------------------------------------------------------------
// 3. OUTPUTS
//------------------------------------------------------------------------------
	//--- COM : control mode status to SCADA, HMI and WEBVISU
	COM.SCADA_OUTPUT_LOCAL_FUXA_ACTIVE := INTERN.LOCAL_FUXA;
	COM.SCADA_OUTPUT_LOCAL_HMI_ACTIVE  := INTERN.LOCAL_HMI;
	COM.HMI_OUTPUT_LOCAL_ACTIVE        := INTERN.LOCAL_HMI;
	COM.WEBVISU_OUTPUT_LOCAL_ACTIVE        := INTERN.LOCAL_WEBVISU;
	COM.WEBVISU_OUTPUT_LOCAL_HMI_ACTIVE  := INTERN.LOCAL_HMI;
	COM.WEBVISU_OUTPUT_LOCAL_FUXA_ACTIVE := INTERN.LOCAL_FUXA;

	//--- EXC
	EXC.EXC_OUTPUT_SIGNAL := INTERN.SIGNAL;

	//--- IO
	IO.OUTPUT_CALIBRATION_HIGH := INTERN.CALIB_HIGH;
	IO.OUTPUT_CALIBRATION_LOW  := INTERN.CALIB_LOW;

	//--- COM : feedback to SCADA, HMI and WEBVISU
	COM.SCADA_OUTPUT_SIGNAL.Real_value := INTERN.SIGNAL;
	COM.HMI_OUTPUT_SIGNAL.Real_value   := INTERN.SIGNAL;
	COM.WEBVISU_OUTPUT_SIGNAL.Real_value   := INTERN.SIGNAL;
	COM.SCADA_OUTPUT_FAULT             := INTERN.FAULT;
	COM.HMI_OUTPUT_FAULT               := INTERN.FAULT;
	COM.WEBVISU_OUTPUT_FAULT               := INTERN.FAULT;
	COM.SCADA_OUTPUT_CALIBRATION_DONE  := INTERN.CALIB_DONE;
	COM.HMI_OUTPUT_CALIBRATION_DONE    := INTERN.CALIB_DONE;
	COM.WEBVISU_OUTPUT_CALIBRATION_DONE    := INTERN.CALIB_DONE;


          
END_FUNCTION_BLOCK
